(* CODESYS project Example10_PLC.project

Project tree, tasks and I/O mapping:
  Device : CODESYS Control Win V3, 3S - Smart Software Solutions GmbH, order no. 305021, version 3.5.7.0
    application Application
      libraries: Standard, * (System)
      task MainTask (cyclic, interval t#20ms, priority 1) calls PLC_PRG
      program PLC_PRG [ST]
      global variables GVL
      function block FB_G4LTL [ST]
    Ethernet : Ethernet, 3S - Smart Software Solutions GmbH, version 3.5.7.0
      Modbus_TCP_Master : Modbus TCP Master, 3S - Smart Software Solutions GmbH, version 3.5.6.0
          settings: AutoReconnect = TRUE
        Modbus_TCP_Slave : Modbus TCP Slave, 3S - Smart Software Solutions GmbH, version 3.5.7.0
            settings: Unit-ID = 1; IPAddress = [127, 0, 0, 1]; Channel 0.Function Code = 4; Channel 0.Read Offset = 16#0000; Channel 0.Read Length = 1; Channel 0.Write Offset = 0; Channel 0.Write Length = 0; Channel 0.Cycle Time = 100; Channel 1.Function Code = 4; Channel 1.Read Offset = 16#0001; Channel 1.Read Length = 1; Channel 1.Write Offset = 0; Channel 1.Write Length = 0; Channel 1.Cycle Time = 100; Channel 2.Function Code = 4; Channel 2.Read Offset = 16#0002; Channel 2.Read Length = 1; Channel 2.Write Offset = 0; Channel 2.Write Length = 0; Channel 2.Cycle Time = 100; Channel 3.Function Code = 4; Channel 3.Read Offset = 16#0003; Channel 3.Read Length = 1; Channel 3.Write Offset = 0; Channel 3.Write Length = 0; Channel 3.Cycle Time = 100; Channel 4.Function Code = 4; Channel 4.Read Offset = 16#0004; Channel 4.Read Length = 1; Channel 4.Write Offset = 0; Channel 4.Write Length = 0; Channel 4.Cycle Time = 100; Channel 5.Function Code = 6; Channel 5.Read Offset = 0; Channel 5.Read Length = 0; Channel 5.Write Offset = 16#0000; Channel 5.Write Length = 1; Channel 5.Cycle Time = 100; Channel 6.Function Code = 6; Channel 6.Read Offset = 0;
              Channel 6.Read Length = 0; Channel 6.Write Offset = 16#0002; Channel 6.Write Length = 1; Channel 6.Cycle Time = 100; Channel 7.Function Code = 6; Channel 7.Read Offset = 0; Channel 7.Read Length = 0; Channel 7.Write Offset = 16#0003; Channel 7.Write Length = 1; Channel 7.Cycle Time = 100; Channel 8.Function Code = 6; Channel 8.Read Offset = 0; Channel 8.Read Length = 0; Channel 8.Write Offset = 16#0004; Channel 8.Write Length = 1; Channel 8.Cycle Time = 100; Channel 9.Function Code = 6; Channel 9.Read Offset = 0; Channel 9.Read Length = 0; Channel 9.Write Offset = 16#0001; Channel 9.Write Length = 1; Channel 9.Cycle Time = 100
            input  Application.dIn0 : BOOL  // Channel 0.Channel 0.Bit0
            input  Application.dIn1 : BOOL  // Channel 1.Channel 1.Bit0
            input  Application.dIn2 : BOOL  // Channel 2.Channel 2.Bit0
            input  Application.dIn3 : BOOL  // Channel 3.Channel 3.Bit0
            input  Application.dIn4 : BOOL  // Channel 4.Channel 4.Bit0
            output Application.dOut0 : BOOL  // Channel 5.Channel 5.Bit0
            output Application.dOut2 : BOOL  // Channel 6.Channel 6.Bit0
            output Application.dOut3 : BOOL  // Channel 7.Channel 7.Bit0
            output Application.dOut4 : BOOL  // Channel 8.Channel 8.Bit0
            output Application.dOut1 : BOOL  // Channel 9.Channel 9.Bit0
            unmapped channels: Channel 0, Channel 1, Channel 2, Channel 3, Channel 4, Channel 5, Channel 6, Channel 7, Channel 8, Channel 9
*)

// Device/Application/GVL
VAR_GLOBAL
	
dIn0 : BOOL;
dIn1 : BOOL;
dIn2 : BOOL;
dIn3 : BOOL;
dIn4 : BOOL;

dOut0 : BOOL;
dOut1 : BOOL; 
dOut2 : BOOL; 
dOut3 : BOOL; 
dOut4 : BOOL; 
END_VAR

// Device/Application/PLC_PRG
PROGRAM PLC_PRG


VAR 
	fb: FB_G4LTL;

END_VAR

// Direct looping
// Assign pins (from global variable to function block) 
fb.x0 := dIn0;
fb.x1 := dIn1;
fb.x2 := dIn2;
fb.x3 := dIn3;
fb.x10 := dIn4;

// Assign pins (from function block to global variable)
dOut0 := fb.y0;
dOut1 := fb.y1;
dOut2 := fb.y2;
dOut3 := fb.y3;

// Run the function block
fb();

END_PROGRAM

// Device/Application/FB_G4LTL
FUNCTION_BLOCK FB_G4LTL

   (* Variable definition *)
   VAR_INPUT
      x0	: BOOL;
      x1	: BOOL;
      x2	: BOOL;
      x3	: BOOL;
      x10	: BOOL;
   END_VAR
   VAR_OUTPUT
      y0	: BOOL;
      y1	: BOOL;
      y2	: BOOL;
      y3	: BOOL;
   END_VAR
   VAR
   (* Control logic for y0, y1; the total number of states equals to 13 *)
      cstate23	: LINT := 0;
   (* Control logic for y2, y3; the total number of states equals to 37 *)
      cstate64	: LINT := 0;  
	  
      t0	: TON;
      t0_reset	: BOOL := FALSE;
      t0_up	: BOOL := FALSE;
      t0_start	: BOOL := FALSE;
      t1	: TON;
      t1_reset	: BOOL := FALSE;
      t1_up	: BOOL := FALSE;
      t1_start	: BOOL := FALSE;
	  
      T0_VALUE	: TIME := TIME#3S;
      T1_VALUE	: TIME := TIME#6S;	  
   END_VAR

   (* Constant definition  *)

    (* Control logic for y0, y1*)
CASE cstate23 OF
262:
    IF ((x0 = TRUE) AND  (x1 = FALSE) AND  ( TRUE ) AND  (x10 = TRUE)) OR ((x0 = TRUE) AND  (x1 = TRUE) AND  (x2 = FALSE) AND  (x10 = TRUE)) OR ((x0 = TRUE) AND  (x1 = TRUE) AND  (x2 = TRUE) AND  ( TRUE )) THEN 
        cstate23 := 27; y0 := FALSE; y1 := FALSE;  
    ELSIF ((x0 = FALSE) AND  (x1 = FALSE) AND  ( TRUE ) AND  (x10 = TRUE)) OR ((x0 = FALSE) AND  (x1 = TRUE) AND  (x2 = FALSE) AND  (x10 = TRUE)) OR ((x0 = FALSE) AND  (x1 = TRUE) AND  (x2 = TRUE) AND  ( TRUE )) THEN 
        cstate23 := 20; y0 := FALSE; y1 := FALSE;  
    ELSIF ((x0 = FALSE) AND  (x1 = FALSE) AND  ( TRUE ) AND  (x10 = FALSE)) THEN 
        cstate23 := 20; y0 := TRUE; y1 := FALSE;  
    ELSIF ((x0 = TRUE) AND  (x1 = TRUE) AND  (x2 = FALSE) AND  (x10 = FALSE)) THEN 
        cstate23 := 265; y0 := FALSE; y1 := TRUE;  
    ELSIF ((x0 = TRUE) AND  (x1 = FALSE) AND  ( TRUE ) AND  (x10 = FALSE)) THEN 
        cstate23 := 262; y0 := TRUE; y1 := FALSE;  
    ELSIF ((x0 = FALSE) AND  (x1 = TRUE) AND  (x2 = FALSE) AND  (x10 = FALSE)) THEN 
        cstate23 := 260; y0 := FALSE; y1 := TRUE;  
    END_IF;
669:
    IF ((x0 = TRUE) AND  (x1 = FALSE) AND  ( TRUE ) AND  (x10 = TRUE)) OR ((x0 = TRUE) AND  (x1 = TRUE) AND  (x2 = FALSE) AND  (x10 = TRUE)) OR ((x0 = TRUE) AND  (x1 = TRUE) AND  (x2 = TRUE) AND  ( TRUE )) THEN 
        cstate23 := 27; y0 := FALSE; y1 := FALSE;  
    ELSIF ((x0 = FALSE) AND  (x1 = FALSE) AND  ( TRUE ) AND  (x10 = TRUE)) OR ((x0 = FALSE) AND  (x1 = TRUE) AND  (x2 = FALSE) AND  (x10 = TRUE)) OR ((x0 = FALSE) AND  (x1 = TRUE) AND  (x2 = TRUE) AND  ( TRUE )) THEN 
        cstate23 := 20; y0 := FALSE; y1 := FALSE;  
    ELSIF ((x0 = FALSE) AND  ( TRUE ) AND  (x2 = FALSE) AND  (x10 = FALSE)) THEN 
        cstate23 := 260; y0 := FALSE; y1 := TRUE;  
    ELSIF ((x0 = TRUE) AND  (x1 = TRUE) AND  (x2 = FALSE) AND  (x10 = FALSE)) THEN 
        cstate23 := 265; y0 := FALSE; y1 := TRUE;  
    ELSIF ((x0 = FALSE) AND  (x1 = FALSE) AND  (x2 = TRUE) AND  (x10 = FALSE)) THEN 
        cstate23 := 20; y0 := TRUE; y1 := FALSE;  
    ELSIF ((x0 = TRUE) AND  (x1 = FALSE) AND  (x2 = TRUE) AND  (x10 = FALSE)) THEN 
        cstate23 := 262; y0 := TRUE; y1 := FALSE;  
    ELSIF ((x0 = TRUE) AND  (x1 = FALSE) AND  (x2 = FALSE) AND  (x10 = FALSE)) THEN 
        cstate23 := 669; y0 := TRUE; y1 := TRUE;  
    END_IF;
260:
    IF ((x0 = TRUE) AND  (x1 = FALSE) AND  ( TRUE ) AND  (x10 = TRUE)) OR ((x0 = TRUE) AND  (x1 = TRUE) AND  (x2 = FALSE) AND  (x10 = TRUE)) OR ((x0 = TRUE) AND  (x1 = TRUE) AND  (x2 = TRUE) AND  ( TRUE )) THEN 
        cstate23 := 27; y0 := FALSE; y1 := FALSE;  
    ELSIF ((x0 = FALSE) AND  ( TRUE ) AND  (x2 = FALSE) AND  (x10 = TRUE)) OR ((x0 = FALSE) AND  ( TRUE ) AND  (x2 = TRUE) AND  ( TRUE )) THEN 
        cstate23 := 20; y0 := FALSE; y1 := FALSE;  
    ELSIF ((x0 = FALSE) AND  ( TRUE ) AND  (x2 = FALSE) AND  (x10 = FALSE)) THEN 
        cstate23 := 260; y0 := FALSE; y1 := TRUE;  
    ELSIF ((x0 = TRUE) AND  (x1 = TRUE) AND  (x2 = FALSE) AND  (x10 = FALSE)) THEN 
        cstate23 := 265; y0 := FALSE; y1 := TRUE;  
    ELSIF ((x0 = TRUE) AND  (x1 = FALSE) AND  (x2 = TRUE) AND  (x10 = FALSE)) THEN 
        cstate23 := 262; y0 := TRUE; y1 := FALSE;  
    ELSIF ((x0 = TRUE) AND  (x1 = FALSE) AND  (x2 = FALSE) AND  (x10 = FALSE)) THEN 
        cstate23 := 669; y0 := TRUE; y1 := TRUE;  
    END_IF;
18:
    IF ((x0 = TRUE) AND  ( TRUE ) AND  ( TRUE ) AND  (x10 = TRUE)) THEN 
        cstate23 := 27; y0 := FALSE; y1 := FALSE;  
    ELSIF ((x0 = FALSE) AND  ( TRUE ) AND  ( TRUE ) AND  (x10 = TRUE)) THEN 
        cstate23 := 20; y0 := FALSE; y1 := FALSE;  
    ELSIF ((x0 = FALSE) AND  (x1 = FALSE) AND  ( TRUE ) AND  (x10 = FALSE)) OR ((x0 = FALSE) AND  (x1 = TRUE) AND  (x2 = TRUE) AND  (x10 = FALSE)) THEN 
        cstate23 := 18; y0 := FALSE; y1 := FALSE;  
    ELSIF ((x0 = TRUE) AND  (x1 = TRUE) AND  (x2 = FALSE) AND  (x10 = FALSE)) THEN 
        cstate23 := 31; y0 := FALSE; y1 := TRUE;  
    ELSIF ((x0 = TRUE) AND  (x1 = TRUE) AND  (x2 = TRUE) AND  (x10 = FALSE)) THEN 
        cstate23 := 25; y0 := FALSE; y1 := FALSE;  
    ELSIF ((x0 = TRUE) AND  (x1 = FALSE) AND  ( TRUE ) AND  (x10 = FALSE)) THEN 
        cstate23 := 257; y0 := TRUE; y1 := FALSE;  
    ELSIF ((x0 = FALSE) AND  (x1 = TRUE) AND  (x2 = FALSE) AND  (x10 = FALSE)) THEN 
        cstate23 := 24; y0 := FALSE; y1 := TRUE;  
    END_IF;
24:
    IF ((x0 = TRUE) AND  ( TRUE ) AND  ( TRUE ) AND  (x10 = TRUE)) THEN 
        cstate23 := 27; y0 := FALSE; y1 := FALSE;  
    ELSIF ((x0 = FALSE) AND  ( TRUE ) AND  ( TRUE ) AND  (x10 = TRUE)) THEN 
        cstate23 := 20; y0 := FALSE; y1 := FALSE;  
    ELSIF ((x0 = FALSE) AND  ( TRUE ) AND  (x2 = FALSE) AND  (x10 = FALSE)) THEN 
        cstate23 := 24; y0 := FALSE; y1 := TRUE;  
    ELSIF ((x0 = TRUE) AND  (x1 = TRUE) AND  (x2 = FALSE) AND  (x10 = FALSE)) THEN 
        cstate23 := 31; y0 := FALSE; y1 := TRUE;  
    ELSIF ((x0 = TRUE) AND  (x1 = TRUE) AND  (x2 = TRUE) AND  (x10 = FALSE)) THEN 
        cstate23 := 25; y0 := FALSE; y1 := FALSE;  
    ELSIF ((x0 = FALSE) AND  ( TRUE ) AND  (x2 = TRUE) AND  (x10 = FALSE)) THEN 
        cstate23 := 18; y0 := FALSE; y1 := FALSE;  
    ELSIF ((x0 = TRUE) AND  (x1 = FALSE) AND  (x2 = TRUE) AND  (x10 = FALSE)) THEN 
        cstate23 := 257; y0 := TRUE; y1 := FALSE;  
    ELSIF ((x0 = TRUE) AND  (x1 = FALSE) AND  (x2 = FALSE) AND  (x10 = FALSE)) THEN 
        cstate23 := 279; y0 := TRUE; y1 := TRUE;  
    END_IF;
25:
    IF ((x0 = TRUE) AND  ( TRUE ) AND  ( TRUE ) AND  (x10 = TRUE)) THEN 
        cstate23 := 27; y0 := FALSE; y1 := FALSE;  
    ELSIF ((x0 = FALSE) AND  ( TRUE ) AND  ( TRUE ) AND  (x10 = TRUE)) THEN 
        cstate23 := 20; y0 := FALSE; y1 := FALSE;  
    ELSIF ((x0 = FALSE) AND  (x1 = FALSE) AND  ( TRUE ) AND  (x10 = FALSE)) THEN 
        cstate23 := 18; y0 := TRUE; y1 := FALSE;  
    ELSIF ((x0 = TRUE) AND  (x1 = TRUE) AND  (x2 = FALSE) AND  (x10 = FALSE)) THEN 
        cstate23 := 31; y0 := FALSE; y1 := TRUE;  
    ELSIF ((x0 = TRUE) AND  (x1 = TRUE) AND  (x2 = TRUE) AND  (x10 = FALSE)) THEN 
        cstate23 := 25; y0 := FALSE; y1 := FALSE;  
    ELSIF ((x0 = FALSE) AND  (x1 = TRUE) AND  (x2 = TRUE) AND  (x10 = FALSE)) THEN 
        cstate23 := 18; y0 := FALSE; y1 := FALSE;  
    ELSIF ((x0 = TRUE) AND  (x1 = FALSE) AND  ( TRUE ) AND  (x10 = FALSE)) THEN 
        cstate23 := 25; y0 := TRUE; y1 := FALSE;  
    ELSIF ((x0 = FALSE) AND  (x1 = TRUE) AND  (x2 = FALSE) AND  (x10 = FALSE)) THEN 
        cstate23 := 24; y0 := FALSE; y1 := TRUE;  
    END_IF;
27:
    IF ((x0 = TRUE) AND  (x1 = FALSE) AND  ( TRUE ) AND  (x10 = TRUE)) OR ((x0 = TRUE) AND  (x1 = TRUE) AND  (x2 = FALSE) AND  (x10 = TRUE)) OR ((x0 = TRUE) AND  (x1 = TRUE) AND  (x2 = TRUE) AND  ( TRUE )) THEN 
        cstate23 := 27; y0 := FALSE; y1 := FALSE;  
    ELSIF ((x0 = FALSE) AND  (x1 = FALSE) AND  ( TRUE ) AND  (x10 = TRUE)) OR ((x0 = FALSE) AND  (x1 = TRUE) AND  (x2 = FALSE) AND  (x10 = TRUE)) OR ((x0 = FALSE) AND  (x1 = TRUE) AND  (x2 = TRUE) AND  ( TRUE )) THEN 
        cstate23 := 20; y0 := FALSE; y1 := FALSE;  
    ELSIF ((x0 = FALSE) AND  (x1 = FALSE) AND  ( TRUE ) AND  (x10 = FALSE)) THEN 
        cstate23 := 20; y0 := TRUE; y1 := FALSE;  
    ELSIF ((x0 = TRUE) AND  (x1 = TRUE) AND  (x2 = FALSE) AND  (x10 = FALSE)) THEN 
        cstate23 := 265; y0 := FALSE; y1 := TRUE;  
    ELSIF ((x0 = TRUE) AND  (x1 = FALSE) AND  ( TRUE ) AND  (x10 = FALSE)) THEN 
        cstate23 := 27; y0 := TRUE; y1 := FALSE;  
    ELSIF ((x0 = FALSE) AND  (x1 = TRUE) AND  (x2 = FALSE) AND  (x10 = FALSE)) THEN 
        cstate23 := 260; y0 := FALSE; y1 := TRUE;  
    END_IF;
20:
    IF ((x0 = TRUE) AND  (x1 = FALSE) AND  ( TRUE ) AND  (x10 = TRUE)) OR ((x0 = TRUE) AND  (x1 = TRUE) AND  (x2 = FALSE) AND  (x10 = TRUE)) OR ((x0 = TRUE) AND  (x1 = TRUE) AND  (x2 = TRUE) AND  ( TRUE )) THEN 
        cstate23 := 27; y0 := FALSE; y1 := FALSE;  
    ELSIF ((x0 = FALSE) AND  (x1 = FALSE) AND  ( TRUE ) AND  ( TRUE )) OR ((x0 = FALSE) AND  (x1 = TRUE) AND  (x2 = FALSE) AND  (x10 = TRUE)) OR ((x0 = FALSE) AND  (x1 = TRUE) AND  (x2 = TRUE) AND  ( TRUE )) THEN 
        cstate23 := 20; y0 := FALSE; y1 := FALSE;  
    ELSIF ((x0 = TRUE) AND  (x1 = TRUE) AND  (x2 = FALSE) AND  (x10 = FALSE)) THEN 
        cstate23 := 265; y0 := FALSE; y1 := TRUE;  
    ELSIF ((x0 = TRUE) AND  (x1 = FALSE) AND  ( TRUE ) AND  (x10 = FALSE)) THEN 
        cstate23 := 262; y0 := TRUE; y1 := FALSE;  
    ELSIF ((x0 = FALSE) AND  (x1 = TRUE) AND  (x2 = FALSE) AND  (x10 = FALSE)) THEN 
        cstate23 := 260; y0 := FALSE; y1 := TRUE;  
    END_IF;
0:
    IF ((x0 = TRUE) AND  ( TRUE ) AND  ( TRUE ) AND  (x10 = TRUE)) THEN 
        cstate23 := 27; y0 := FALSE; y1 := FALSE;  
    ELSIF ((x0 = FALSE) AND  ( TRUE ) AND  ( TRUE ) AND  (x10 = TRUE)) THEN 
        cstate23 := 20; y0 := FALSE; y1 := FALSE;  
    ELSIF ((x0 = FALSE) AND  (x1 = FALSE) AND  ( TRUE ) AND  (x10 = FALSE)) OR ((x0 = FALSE) AND  (x1 = TRUE) AND  (x2 = TRUE) AND  (x10 = FALSE)) THEN 
        cstate23 := 18; y0 := FALSE; y1 := FALSE;  
    ELSIF ((x0 = TRUE) AND  (x1 = TRUE) AND  (x2 = FALSE) AND  (x10 = FALSE)) THEN 
        cstate23 := 31; y0 := FALSE; y1 := TRUE;  
    ELSIF ((x0 = TRUE) AND  (x1 = FALSE) AND  ( TRUE ) AND  (x10 = FALSE)) OR ((x0 = TRUE) AND  (x1 = TRUE) AND  (x2 = TRUE) AND  (x10 = FALSE)) THEN 
        cstate23 := 25; y0 := FALSE; y1 := FALSE;  
    ELSIF ((x0 = FALSE) AND  (x1 = TRUE) AND  (x2 = FALSE) AND  (x10 = FALSE)) THEN 
        cstate23 := 24; y0 := FALSE; y1 := TRUE;  
    END_IF;
279:
    IF ((x0 = TRUE) AND  ( TRUE ) AND  ( TRUE ) AND  (x10 = TRUE)) THEN 
        cstate23 := 27; y0 := FALSE; y1 := FALSE;  
    ELSIF ((x0 = FALSE) AND  ( TRUE ) AND  ( TRUE ) AND  (x10 = TRUE)) THEN 
        cstate23 := 20; y0 := FALSE; y1 := FALSE;  
    ELSIF ((x0 = FALSE) AND  ( TRUE ) AND  (x2 = FALSE) AND  (x10 = FALSE)) THEN 
        cstate23 := 24; y0 := FALSE; y1 := TRUE;  
    ELSIF ((x0 = TRUE) AND  (x1 = TRUE) AND  (x2 = FALSE) AND  (x10 = FALSE)) THEN 
        cstate23 := 31; y0 := FALSE; y1 := TRUE;  
    ELSIF ((x0 = TRUE) AND  (x1 = TRUE) AND  (x2 = TRUE) AND  (x10 = FALSE)) THEN 
        cstate23 := 25; y0 := FALSE; y1 := FALSE;  
    ELSIF ((x0 = FALSE) AND  (x1 = FALSE) AND  (x2 = TRUE) AND  (x10 = FALSE)) THEN 
        cstate23 := 18; y0 := TRUE; y1 := FALSE;  
    ELSIF ((x0 = FALSE) AND  (x1 = TRUE) AND  (x2 = TRUE) AND  (x10 = FALSE)) THEN 
        cstate23 := 18; y0 := FALSE; y1 := FALSE;  
    ELSIF ((x0 = TRUE) AND  (x1 = FALSE) AND  (x2 = TRUE) AND  (x10 = FALSE)) THEN 
        cstate23 := 257; y0 := TRUE; y1 := FALSE;  
    ELSIF ((x0 = TRUE) AND  (x1 = FALSE) AND  (x2 = FALSE) AND  (x10 = FALSE)) THEN 
        cstate23 := 279; y0 := TRUE; y1 := TRUE;  
    END_IF;
31:
    IF ((x0 = TRUE) AND  ( TRUE ) AND  ( TRUE ) AND  (x10 = TRUE)) THEN 
        cstate23 := 27; y0 := FALSE; y1 := FALSE;  
    ELSIF ((x0 = FALSE) AND  ( TRUE ) AND  ( TRUE ) AND  (x10 = TRUE)) THEN 
        cstate23 := 20; y0 := FALSE; y1 := FALSE;  
    ELSIF ((x0 = FALSE) AND  ( TRUE ) AND  (x2 = FALSE) AND  (x10 = FALSE)) THEN 
        cstate23 := 24; y0 := FALSE; y1 := TRUE;  
    ELSIF ((x0 = TRUE) AND  ( TRUE ) AND  (x2 = FALSE) AND  (x10 = FALSE)) THEN 
        cstate23 := 31; y0 := FALSE; y1 := TRUE;  
    ELSIF ((x0 = TRUE) AND  (x1 = TRUE) AND  (x2 = TRUE) AND  (x10 = FALSE)) THEN 
        cstate23 := 25; y0 := FALSE; y1 := FALSE;  
    ELSIF ((x0 = FALSE) AND  (x1 = FALSE) AND  (x2 = TRUE) AND  (x10 = FALSE)) THEN 
        cstate23 := 18; y0 := TRUE; y1 := FALSE;  
    ELSIF ((x0 = FALSE) AND  (x1 = TRUE) AND  (x2 = TRUE) AND  (x10 = FALSE)) THEN 
        cstate23 := 18; y0 := FALSE; y1 := FALSE;  
    ELSIF ((x0 = TRUE) AND  (x1 = FALSE) AND  (x2 = TRUE) AND  (x10 = FALSE)) THEN 
        cstate23 := 25; y0 := TRUE; y1 := FALSE;  
    END_IF;
257:
    IF ((x0 = TRUE) AND  ( TRUE ) AND  ( TRUE ) AND  (x10 = TRUE)) THEN 
        cstate23 := 27; y0 := FALSE; y1 := FALSE;  
    ELSIF ((x0 = FALSE) AND  ( TRUE ) AND  ( TRUE ) AND  (x10 = TRUE)) THEN 
        cstate23 := 20; y0 := FALSE; y1 := FALSE;  
    ELSIF ((x0 = FALSE) AND  (x1 = FALSE) AND  ( TRUE ) AND  (x10 = FALSE)) THEN 
        cstate23 := 18; y0 := TRUE; y1 := FALSE;  
    ELSIF ((x0 = TRUE) AND  (x1 = TRUE) AND  (x2 = FALSE) AND  (x10 = FALSE)) THEN 
        cstate23 := 31; y0 := FALSE; y1 := TRUE;  
    ELSIF ((x0 = TRUE) AND  (x1 = TRUE) AND  (x2 = TRUE) AND  (x10 = FALSE)) THEN 
        cstate23 := 25; y0 := FALSE; y1 := FALSE;  
    ELSIF ((x0 = FALSE) AND  (x1 = TRUE) AND  (x2 = TRUE) AND  (x10 = FALSE)) THEN 
        cstate23 := 18; y0 := FALSE; y1 := FALSE;  
    ELSIF ((x0 = TRUE) AND  (x1 = FALSE) AND  ( TRUE ) AND  (x10 = FALSE)) THEN 
        cstate23 := 257; y0 := TRUE; y1 := FALSE;  
    ELSIF ((x0 = FALSE) AND  (x1 = TRUE) AND  (x2 = FALSE) AND  (x10 = FALSE)) THEN 
        cstate23 := 24; y0 := FALSE; y1 := TRUE;  
    END_IF;
265:
    IF ((x0 = TRUE) AND  (x1 = FALSE) AND  ( TRUE ) AND  (x10 = TRUE)) OR ((x0 = TRUE) AND  (x1 = TRUE) AND  (x2 = FALSE) AND  (x10 = TRUE)) OR ((x0 = TRUE) AND  (x1 = TRUE) AND  (x2 = TRUE) AND  ( TRUE )) THEN 
        cstate23 := 27; y0 := FALSE; y1 := FALSE;  
    ELSIF ((x0 = FALSE) AND  (x1 = FALSE) AND  ( TRUE ) AND  (x10 = TRUE)) OR ((x0 = FALSE) AND  (x1 = TRUE) AND  (x2 = FALSE) AND  (x10 = TRUE)) OR ((x0 = FALSE) AND  (x1 = TRUE) AND  (x2 = TRUE) AND  ( TRUE )) THEN 
        cstate23 := 20; y0 := FALSE; y1 := FALSE;  
    ELSIF ((x0 = FALSE) AND  ( TRUE ) AND  (x2 = FALSE) AND  (x10 = FALSE)) THEN 
        cstate23 := 260; y0 := FALSE; y1 := TRUE;  
    ELSIF ((x0 = TRUE) AND  ( TRUE ) AND  (x2 = FALSE) AND  (x10 = FALSE)) THEN 
        cstate23 := 265; y0 := FALSE; y1 := TRUE;  
    ELSIF ((x0 = FALSE) AND  (x1 = FALSE) AND  (x2 = TRUE) AND  (x10 = FALSE)) THEN 
        cstate23 := 20; y0 := TRUE; y1 := FALSE;  
    ELSIF ((x0 = TRUE) AND  (x1 = FALSE) AND  (x2 = TRUE) AND  (x10 = FALSE)) THEN 
        cstate23 := 27; y0 := TRUE; y1 := FALSE;  
    END_IF;
END_CASE;


 (* Control logic *)
CASE cstate64 OF
19:
    IF ((x2 = FALSE) AND  ( TRUE ) AND  ( TRUE ) AND  (t0.Q = FALSE) AND  (t1.Q = FALSE)) THEN 
        cstate64 := 19; y2 := FALSE; y3 := FALSE; t0_start := FALSE;t1_start := FALSE; 
    ELSIF ((x2 = FALSE) AND  ( TRUE ) AND  (x10 = FALSE) AND  (t0.Q = FALSE) AND  (t1.Q = TRUE)) THEN 
        cstate64 := 20; y2 := FALSE; y3 := FALSE; t0_start := FALSE;t1_start := FALSE; 
    ELSIF ((x2 = FALSE) AND  ( TRUE ) AND  (x10 = FALSE) AND  (t0.Q = TRUE) AND  ( TRUE )) THEN 
        cstate64 := 37; y2 := FALSE; y3 := TRUE; t0_start := FALSE;t1_start := TRUE; t1_up := FALSE; 
    ELSIF ((x2 = FALSE) AND  ( TRUE ) AND  (x10 = TRUE) AND  (t0.Q = FALSE) AND  (t1.Q = TRUE)) THEN 
        cstate64 := 20; y2 := FALSE; y3 := FALSE; t0_start := FALSE;t1_start := FALSE; 
    ELSIF ((x2 = FALSE) AND  ( TRUE ) AND  (x10 = TRUE) AND  (t0.Q = TRUE) AND  (t1.Q = FALSE)) THEN 
        cstate64 := 34; y2 := FALSE; y3 := FALSE; t0_start := FALSE;t1_start := FALSE; 
    ELSIF ((x2 = FALSE) AND  ( TRUE ) AND  (x10 = TRUE) AND  (t0.Q = TRUE) AND  (t1.Q = TRUE)) THEN 
        cstate64 := 33; y2 := FALSE; y3 := FALSE; t0_start := FALSE;t1_start := FALSE; 
    ELSIF ((x2 = TRUE) AND  ( TRUE ) AND  (x10 = FALSE) AND  (t0.Q = FALSE) AND  (t1.Q = FALSE)) THEN 
        cstate64 := 83; y2 := TRUE; y3 := FALSE; t0_start := TRUE; t0_up := FALSE;t1_start := FALSE; 
    ELSIF ((x2 = TRUE) AND  ( TRUE ) AND  (x10 = FALSE) AND  (t0.Q = FALSE) AND  (t1.Q = TRUE)) THEN 
        cstate64 := 84; y2 := TRUE; y3 := FALSE; t0_start := TRUE; t0_up := FALSE;t1_start := FALSE; 
    ELSIF ((x2 = TRUE) AND  ( TRUE ) AND  (x10 = FALSE) AND  (t0.Q = TRUE) AND  ( TRUE )) THEN 
        cstate64 := 86; y2 := TRUE; y3 := TRUE; t0_start := TRUE; t0_up := FALSE;t1_start := TRUE; t1_up := FALSE; 
    ELSIF ((x2 = TRUE) AND  ( TRUE ) AND  (x10 = TRUE) AND  (t0.Q = FALSE) AND  (t1.Q = FALSE)) THEN 
        cstate64 := 51; y2 := FALSE; y3 := FALSE; t0_start := FALSE;t1_start := FALSE; 
    ELSIF ((x2 = TRUE) AND  ( TRUE ) AND  (x10 = TRUE) AND  (t0.Q = FALSE) AND  (t1.Q = TRUE)) THEN 
        cstate64 := 52; y2 := FALSE; y3 := FALSE; t0_start := FALSE;t1_start := FALSE; 
    ELSIF ((x2 = TRUE) AND  ( TRUE ) AND  (x10 = TRUE) AND  (t0.Q = TRUE) AND  (t1.Q = FALSE)) THEN 
        cstate64 := 66; y2 := FALSE; y3 := FALSE; t0_start := FALSE;t1_start := FALSE; 
    ELSIF ((x2 = TRUE) AND  ( TRUE ) AND  (x10 = TRUE) AND  (t0.Q = TRUE) AND  (t1.Q = TRUE)) THEN 
        cstate64 := 65; y2 := FALSE; y3 := FALSE; t0_start := FALSE;t1_start := FALSE; 
    END_IF;
35:
    IF ((x2 = FALSE) AND  ( TRUE ) AND  ( TRUE ) AND  (t0.Q = FALSE) AND  (t1.Q = FALSE)) THEN 
        cstate64 := 35; y2 := FALSE; y3 := FALSE; t0_start := FALSE;t1_start := FALSE; 
    ELSIF ((x2 = FALSE) AND  ( TRUE ) AND  (x10 = FALSE) AND  (t0.Q = FALSE) AND  (t1.Q = TRUE)) THEN 
        cstate64 := 36; y2 := FALSE; y3 := FALSE; t0_start := FALSE;t1_start := FALSE; 
    ELSIF ((x2 = FALSE) AND  ( TRUE ) AND  (x10 = FALSE) AND  (t0.Q = TRUE) AND  ( TRUE )) THEN 
        cstate64 := 37; y2 := FALSE; y3 := TRUE; t0_start := FALSE;t1_start := TRUE; t1_up := FALSE; 
    ELSIF ((x2 = FALSE) AND  ( TRUE ) AND  (x10 = TRUE) AND  (t0.Q = FALSE) AND  (t1.Q = TRUE)) THEN 
        cstate64 := 36; y2 := FALSE; y3 := FALSE; t0_start := FALSE;t1_start := FALSE; 
    ELSIF ((x2 = FALSE) AND  ( TRUE ) AND  (x10 = TRUE) AND  (t0.Q = TRUE) AND  (t1.Q = FALSE)) THEN 
        cstate64 := 34; y2 := FALSE; y3 := FALSE; t0_start := FALSE;t1_start := FALSE; 
    ELSIF ((x2 = FALSE) AND  ( TRUE ) AND  (x10 = TRUE) AND  (t0.Q = TRUE) AND  (t1.Q = TRUE)) THEN 
        cstate64 := 33; y2 := FALSE; y3 := FALSE; t0_start := FALSE;t1_start := FALSE; 
    ELSIF ((x2 = TRUE) AND  ( TRUE ) AND  (x10 = FALSE) AND  (t0.Q = FALSE) AND  (t1.Q = FALSE)) THEN 
        cstate64 := 83; y2 := TRUE; y3 := FALSE; t0_start := TRUE; t0_up := FALSE;t1_start := FALSE; 
    ELSIF ((x2 = TRUE) AND  ( TRUE ) AND  (x10 = FALSE) AND  (t0.Q = FALSE) AND  (t1.Q = TRUE)) THEN 
        cstate64 := 84; y2 := TRUE; y3 := FALSE; t0_start := TRUE; t0_up := FALSE;t1_start := FALSE; 
    ELSIF ((x2 = TRUE) AND  ( TRUE ) AND  (x10 = FALSE) AND  (t0.Q = TRUE) AND  ( TRUE )) THEN 
        cstate64 := 86; y2 := TRUE; y3 := TRUE; t0_start := TRUE; t0_up := FALSE;t1_start := TRUE; t1_up := FALSE; 
    ELSIF ((x2 = TRUE) AND  ( TRUE ) AND  (x10 = TRUE) AND  (t0.Q = FALSE) AND  (t1.Q = FALSE)) THEN 
        cstate64 := 67; y2 := FALSE; y3 := FALSE; t0_start := FALSE;t1_start := FALSE; 
    ELSIF ((x2 = TRUE) AND  ( TRUE ) AND  (x10 = TRUE) AND  (t0.Q = FALSE) AND  (t1.Q = TRUE)) THEN 
        cstate64 := 68; y2 := FALSE; y3 := FALSE; t0_start := FALSE;t1_start := FALSE; 
    ELSIF ((x2 = TRUE) AND  ( TRUE ) AND  (x10 = TRUE) AND  (t0.Q = TRUE) AND  (t1.Q = FALSE)) THEN 
        cstate64 := 66; y2 := FALSE; y3 := FALSE; t0_start := FALSE;t1_start := FALSE; 
    ELSIF ((x2 = TRUE) AND  ( TRUE ) AND  (x10 = TRUE) AND  (t0.Q = TRUE) AND  (t1.Q = TRUE)) THEN 
        cstate64 := 65; y2 := FALSE; y3 := FALSE; t0_start := FALSE;t1_start := FALSE; 
    END_IF;
36:
    IF ((x2 = FALSE) AND  ( TRUE ) AND  (x10 = FALSE) AND  (t0.Q = FALSE) AND  (t1.Q = FALSE)) OR ((x2 = FALSE) AND  ( TRUE ) AND  (x10 = TRUE) AND  (t0.Q = FALSE) AND  ( TRUE )) THEN 
        cstate64 := 36; y2 := FALSE; y3 := FALSE; t0_start := FALSE;t1_start := FALSE; 
    ELSIF ((x2 = FALSE) AND  ( TRUE ) AND  (x10 = FALSE) AND  (t0.Q = FALSE) AND  (t1.Q = TRUE)) THEN 
        cstate64 := 36; y2 := FALSE; y3 := FALSE; t0_start := FALSE;t1_start := FALSE; 
    ELSIF ((x2 = FALSE) AND  ( TRUE ) AND  (x10 = FALSE) AND  (t0.Q = TRUE) AND  ( TRUE )) THEN 
        cstate64 := 40; y2 := FALSE; y3 := TRUE; t0_start := FALSE;t1_start := TRUE; t1_up := FALSE; 
    ELSIF ((x2 = FALSE) AND  ( TRUE ) AND  (x10 = TRUE) AND  (t0.Q = TRUE) AND  ( TRUE )) THEN 
        cstate64 := 33; y2 := FALSE; y3 := FALSE; t0_start := FALSE;t1_start := FALSE; 
    ELSIF ((x2 = TRUE) AND  ( TRUE ) AND  (x10 = FALSE) AND  (t0.Q = FALSE) AND  (t1.Q = FALSE)) THEN 
        cstate64 := 84; y2 := TRUE; y3 := FALSE; t0_start := TRUE; t0_up := FALSE;t1_start := FALSE; 
    ELSIF ((x2 = TRUE) AND  ( TRUE ) AND  (x10 = FALSE) AND  (t0.Q = FALSE) AND  (t1.Q = TRUE)) THEN 
        cstate64 := 84; y2 := TRUE; y3 := FALSE; t0_start := TRUE; t0_up := FALSE;t1_start := FALSE; 
    ELSIF ((x2 = TRUE) AND  ( TRUE ) AND  (x10 = FALSE) AND  (t0.Q = TRUE) AND  ( TRUE )) THEN 
        cstate64 := 87; y2 := TRUE; y3 := TRUE; t0_start := TRUE; t0_up := FALSE;t1_start := TRUE; t1_up := FALSE; 
    ELSIF ((x2 = TRUE) AND  ( TRUE ) AND  (x10 = TRUE) AND  (t0.Q = FALSE) AND  ( TRUE )) THEN 
        cstate64 := 68; y2 := FALSE; y3 := FALSE; t0_start := FALSE;t1_start := FALSE; 
    ELSIF ((x2 = TRUE) AND  ( TRUE ) AND  (x10 = TRUE) AND  (t0.Q = TRUE) AND  ( TRUE )) THEN 
        cstate64 := 65; y2 := FALSE; y3 := FALSE; t0_start := FALSE;t1_start := FALSE; 
    END_IF;
33:
    IF ((x2 = FALSE) AND  ( TRUE ) AND  (x10 = FALSE) AND  (t0.Q = FALSE) AND  (t1.Q = FALSE)) OR ((x2 = FALSE) AND  ( TRUE ) AND  (x10 = TRUE) AND  (t0.Q = FALSE) AND  ( TRUE )) THEN 
        cstate64 := 36; y2 := FALSE; y3 := FALSE; t0_start := FALSE;t1_start := FALSE; 
    ELSIF ((x2 = FALSE) AND  ( TRUE ) AND  (x10 = FALSE) AND  (t0.Q = FALSE) AND  (t1.Q = TRUE)) THEN 
        cstate64 := 36; y2 := FALSE; y3 := FALSE; t0_start := FALSE;t1_start := FALSE; 
    ELSIF ((x2 = FALSE) AND  ( TRUE ) AND  (x10 = FALSE) AND  (t0.Q = TRUE) AND  ( TRUE )) THEN 
        cstate64 := 33; y2 := FALSE; y3 := FALSE; t0_start := FALSE;t1_start := FALSE; 
    ELSIF ((x2 = FALSE) AND  ( TRUE ) AND  (x10 = TRUE) AND  (t0.Q = TRUE) AND  ( TRUE )) THEN 
        cstate64 := 33; y2 := FALSE; y3 := FALSE; t0_start := FALSE;t1_start := FALSE; 
    ELSIF ((x2 = TRUE) AND  ( TRUE ) AND  (x10 = FALSE) AND  (t0.Q = FALSE) AND  (t1.Q = FALSE)) THEN 
        cstate64 := 84; y2 := TRUE; y3 := FALSE; t0_start := TRUE; t0_up := FALSE;t1_start := FALSE; 
    ELSIF ((x2 = TRUE) AND  ( TRUE ) AND  (x10 = FALSE) AND  (t0.Q = FALSE) AND  (t1.Q = TRUE)) THEN 
        cstate64 := 84; y2 := TRUE; y3 := FALSE; t0_start := TRUE; t0_up := FALSE;t1_start := FALSE; 
    ELSIF ((x2 = TRUE) AND  ( TRUE ) AND  (x10 = FALSE) AND  (t0.Q = TRUE) AND  ( TRUE )) THEN 
        cstate64 := 81; y2 := TRUE; y3 := FALSE; t0_start := TRUE; t0_up := FALSE;t1_start := FALSE; 
    ELSIF ((x2 = TRUE) AND  ( TRUE ) AND  (x10 = TRUE) AND  (t0.Q = FALSE) AND  ( TRUE )) THEN 
        cstate64 := 68; y2 := FALSE; y3 := FALSE; t0_start := FALSE;t1_start := FALSE; 
    ELSIF ((x2 = TRUE) AND  ( TRUE ) AND  (x10 = TRUE) AND  (t0.Q = TRUE) AND  ( TRUE )) THEN 
        cstate64 := 65; y2 := FALSE; y3 := FALSE; t0_start := FALSE;t1_start := FALSE; 
    END_IF;
34:
    IF ((x2 = FALSE) AND  ( TRUE ) AND  ( TRUE ) AND  (t0.Q = FALSE) AND  (t1.Q = FALSE)) THEN 
        cstate64 := 35; y2 := FALSE; y3 := FALSE; t0_start := FALSE;t1_start := FALSE; 
    ELSIF ((x2 = FALSE) AND  ( TRUE ) AND  (x10 = FALSE) AND  (t0.Q = FALSE) AND  (t1.Q = TRUE)) THEN 
        cstate64 := 36; y2 := FALSE; y3 := FALSE; t0_start := FALSE;t1_start := FALSE; 
    ELSIF ((x2 = FALSE) AND  ( TRUE ) AND  (x10 = FALSE) AND  (t0.Q = TRUE) AND  (t1.Q = FALSE)) THEN 
        cstate64 := 34; y2 := FALSE; y3 := FALSE; t0_start := FALSE;t1_start := FALSE; 
    ELSIF ((x2 = FALSE) AND  ( TRUE ) AND  (x10 = FALSE) AND  (t0.Q = TRUE) AND  (t1.Q = TRUE)) THEN 
        cstate64 := 33; y2 := FALSE; y3 := FALSE; t0_start := FALSE;t1_start := FALSE; 
    ELSIF ((x2 = FALSE) AND  ( TRUE ) AND  (x10 = TRUE) AND  (t0.Q = FALSE) AND  (t1.Q = TRUE)) THEN 
        cstate64 := 36; y2 := FALSE; y3 := FALSE; t0_start := FALSE;t1_start := FALSE; 
    ELSIF ((x2 = FALSE) AND  ( TRUE ) AND  (x10 = TRUE) AND  (t0.Q = TRUE) AND  (t1.Q = FALSE)) THEN 
        cstate64 := 34; y2 := FALSE; y3 := FALSE; t0_start := FALSE;t1_start := FALSE; 
    ELSIF ((x2 = FALSE) AND  ( TRUE ) AND  (x10 = TRUE) AND  (t0.Q = TRUE) AND  (t1.Q = TRUE)) THEN 
        cstate64 := 33; y2 := FALSE; y3 := FALSE; t0_start := FALSE;t1_start := FALSE; 
    ELSIF ((x2 = TRUE) AND  ( TRUE ) AND  (x10 = FALSE) AND  (t0.Q = FALSE) AND  (t1.Q = FALSE)) THEN 
        cstate64 := 83; y2 := TRUE; y3 := FALSE; t0_start := TRUE; t0_up := FALSE;t1_start := FALSE; 
    ELSIF ((x2 = TRUE) AND  ( TRUE ) AND  (x10 = FALSE) AND  (t0.Q = FALSE) AND  (t1.Q = TRUE)) THEN 
        cstate64 := 84; y2 := TRUE; y3 := FALSE; t0_start := TRUE; t0_up := FALSE;t1_start := FALSE; 
    ELSIF ((x2 = TRUE) AND  ( TRUE ) AND  (x10 = FALSE) AND  (t0.Q = TRUE) AND  (t1.Q = FALSE)) THEN 
        cstate64 := 82; y2 := TRUE; y3 := FALSE; t0_start := TRUE; t0_up := FALSE;t1_start := FALSE; 
    ELSIF ((x2 = TRUE) AND  ( TRUE ) AND  (x10 = FALSE) AND  (t0.Q = TRUE) AND  (t1.Q = TRUE)) THEN 
        cstate64 := 81; y2 := TRUE; y3 := FALSE; t0_start := TRUE; t0_up := FALSE;t1_start := FALSE; 
    ELSIF ((x2 = TRUE) AND  ( TRUE ) AND  (x10 = TRUE) AND  (t0.Q = FALSE) AND  (t1.Q = FALSE)) THEN 
        cstate64 := 67; y2 := FALSE; y3 := FALSE; t0_start := FALSE;t1_start := FALSE; 
    ELSIF ((x2 = TRUE) AND  ( TRUE ) AND  (x10 = TRUE) AND  (t0.Q = FALSE) AND  (t1.Q = TRUE)) THEN 
        cstate64 := 68; y2 := FALSE; y3 := FALSE; t0_start := FALSE;t1_start := FALSE; 
    ELSIF ((x2 = TRUE) AND  ( TRUE ) AND  (x10 = TRUE) AND  (t0.Q = TRUE) AND  (t1.Q = FALSE)) THEN 
        cstate64 := 66; y2 := FALSE; y3 := FALSE; t0_start := FALSE;t1_start := FALSE; 
    ELSIF ((x2 = TRUE) AND  ( TRUE ) AND  (x10 = TRUE) AND  (t0.Q = TRUE) AND  (t1.Q = TRUE)) THEN 
        cstate64 := 65; y2 := FALSE; y3 := FALSE; t0_start := FALSE;t1_start := FALSE; 
    END_IF;
37:
    IF ((x2 = FALSE) AND  ( TRUE ) AND  (x10 = FALSE) AND  (t0.Q = FALSE) AND  (t1.Q = FALSE)) THEN 
        cstate64 := 41; y2 := FALSE; y3 := TRUE; t0_start := FALSE;t1_start := FALSE; 
    ELSIF ((x2 = FALSE) AND  ( TRUE ) AND  (x10 = FALSE) AND  (t0.Q = FALSE) AND  (t1.Q = TRUE)) THEN 
        cstate64 := 36; y2 := FALSE; y3 := FALSE; t0_start := FALSE;t1_start := FALSE; 
    ELSIF ((x2 = FALSE) AND  ( TRUE ) AND  (x10 = FALSE) AND  (t0.Q = TRUE) AND  (t1.Q = FALSE)) THEN 
        cstate64 := 37; y2 := FALSE; y3 := TRUE; t0_start := FALSE;t1_start := FALSE; 
    ELSIF ((x2 = FALSE) AND  ( TRUE ) AND  (x10 = FALSE) AND  (t0.Q = TRUE) AND  (t1.Q = TRUE)) THEN 
        cstate64 := 33; y2 := FALSE; y3 := FALSE; t0_start := FALSE;t1_start := FALSE; 
    ELSIF ((x2 = FALSE) AND  ( TRUE ) AND  (x10 = TRUE) AND  (t0.Q = FALSE) AND  (t1.Q = FALSE)) THEN 
        cstate64 := 35; y2 := FALSE; y3 := FALSE; t0_start := FALSE;t1_start := FALSE; 
    ELSIF ((x2 = FALSE) AND  ( TRUE ) AND  (x10 = TRUE) AND  (t0.Q = FALSE) AND  (t1.Q = TRUE)) THEN 
        cstate64 := 36; y2 := FALSE; y3 := FALSE; t0_start := FALSE;t1_start := FALSE; 
    ELSIF ((x2 = FALSE) AND  ( TRUE ) AND  (x10 = TRUE) AND  (t0.Q = TRUE) AND  (t1.Q = FALSE)) THEN 
        cstate64 := 34; y2 := FALSE; y3 := FALSE; t0_start := FALSE;t1_start := FALSE; 
    ELSIF ((x2 = FALSE) AND  ( TRUE ) AND  (x10 = TRUE) AND  (t0.Q = TRUE) AND  (t1.Q = TRUE)) THEN 
        cstate64 := 33; y2 := FALSE; y3 := FALSE; t0_start := FALSE;t1_start := FALSE; 
    ELSIF ((x2 = TRUE) AND  ( TRUE ) AND  (x10 = FALSE) AND  (t0.Q = FALSE) AND  (t1.Q = FALSE)) THEN 
        cstate64 := 90; y2 := TRUE; y3 := TRUE; t0_start := TRUE; t0_up := FALSE;t1_start := FALSE; 
    ELSIF ((x2 = TRUE) AND  ( TRUE ) AND  (x10 = FALSE) AND  (t0.Q = FALSE) AND  (t1.Q = TRUE)) THEN 
        cstate64 := 84; y2 := TRUE; y3 := FALSE; t0_start := TRUE; t0_up := FALSE;t1_start := FALSE; 
    ELSIF ((x2 = TRUE) AND  ( TRUE ) AND  (x10 = FALSE) AND  (t0.Q = TRUE) AND  (t1.Q = FALSE)) THEN 
        cstate64 := 86; y2 := TRUE; y3 := TRUE; t0_start := TRUE; t0_up := FALSE;t1_start := FALSE; 
    ELSIF ((x2 = TRUE) AND  ( TRUE ) AND  (x10 = FALSE) AND  (t0.Q = TRUE) AND  (t1.Q = TRUE)) THEN 
        cstate64 := 81; y2 := TRUE; y3 := FALSE; t0_start := TRUE; t0_up := FALSE;t1_start := FALSE; 
    ELSIF ((x2 = TRUE) AND  ( TRUE ) AND  (x10 = TRUE) AND  (t0.Q = FALSE) AND  (t1.Q = FALSE)) THEN 
        cstate64 := 67; y2 := FALSE; y3 := FALSE; t0_start := FALSE;t1_start := FALSE; 
    ELSIF ((x2 = TRUE) AND  ( TRUE ) AND  (x10 = TRUE) AND  (t0.Q = FALSE) AND  (t1.Q = TRUE)) THEN 
        cstate64 := 68; y2 := FALSE; y3 := FALSE; t0_start := FALSE;t1_start := FALSE; 
    ELSIF ((x2 = TRUE) AND  ( TRUE ) AND  (x10 = TRUE) AND  (t0.Q = TRUE) AND  (t1.Q = FALSE)) THEN 
        cstate64 := 66; y2 := FALSE; y3 := FALSE; t0_start := FALSE;t1_start := FALSE; 
    ELSIF ((x2 = TRUE) AND  ( TRUE ) AND  (x10 = TRUE) AND  (t0.Q = TRUE) AND  (t1.Q = TRUE)) THEN 
        cstate64 := 65; y2 := FALSE; y3 := FALSE; t0_start := FALSE;t1_start := FALSE; 
    END_IF;
20:
    IF ((x2 = FALSE) AND  ( TRUE ) AND  (x10 = FALSE) AND  (t0.Q = FALSE) AND  (t1.Q = FALSE)) OR ((x2 = FALSE) AND  ( TRUE ) AND  (x10 = TRUE) AND  (t0.Q = FALSE) AND  ( TRUE )) THEN 
        cstate64 := 20; y2 := FALSE; y3 := FALSE; t0_start := FALSE;t1_start := FALSE; 
    ELSIF ((x2 = FALSE) AND  ( TRUE ) AND  (x10 = FALSE) AND  (t0.Q = FALSE) AND  (t1.Q = TRUE)) THEN 
        cstate64 := 20; y2 := FALSE; y3 := FALSE; t0_start := FALSE;t1_start := FALSE; 
    ELSIF ((x2 = FALSE) AND  ( TRUE ) AND  (x10 = FALSE) AND  (t0.Q = TRUE) AND  ( TRUE )) THEN 
        cstate64 := 40; y2 := FALSE; y3 := TRUE; t0_start := FALSE;t1_start := TRUE; t1_up := FALSE; 
    ELSIF ((x2 = FALSE) AND  ( TRUE ) AND  (x10 = TRUE) AND  (t0.Q = TRUE) AND  ( TRUE )) THEN 
        cstate64 := 33; y2 := FALSE; y3 := FALSE; t0_start := FALSE;t1_start := FALSE; 
    ELSIF ((x2 = TRUE) AND  ( TRUE ) AND  (x10 = FALSE) AND  (t0.Q = FALSE) AND  (t1.Q = FALSE)) THEN 
        cstate64 := 84; y2 := TRUE; y3 := FALSE; t0_start := TRUE; t0_up := FALSE;t1_start := FALSE; 
    ELSIF ((x2 = TRUE) AND  ( TRUE ) AND  (x10 = FALSE) AND  (t0.Q = FALSE) AND  (t1.Q = TRUE)) THEN 
        cstate64 := 84; y2 := TRUE; y3 := FALSE; t0_start := TRUE; t0_up := FALSE;t1_start := FALSE; 
    ELSIF ((x2 = TRUE) AND  ( TRUE ) AND  (x10 = FALSE) AND  (t0.Q = TRUE) AND  ( TRUE )) THEN 
        cstate64 := 87; y2 := TRUE; y3 := TRUE; t0_start := TRUE; t0_up := FALSE;t1_start := TRUE; t1_up := FALSE; 
    ELSIF ((x2 = TRUE) AND  ( TRUE ) AND  (x10 = TRUE) AND  (t0.Q = FALSE) AND  ( TRUE )) THEN 
        cstate64 := 52; y2 := FALSE; y3 := FALSE; t0_start := FALSE;t1_start := FALSE; 
    ELSIF ((x2 = TRUE) AND  ( TRUE ) AND  (x10 = TRUE) AND  (t0.Q = TRUE) AND  ( TRUE )) THEN 
        cstate64 := 65; y2 := FALSE; y3 := FALSE; t0_start := FALSE;t1_start := FALSE; 
    END_IF;
41:
    IF ((x2 = FALSE) AND  ( TRUE ) AND  (x10 = FALSE) AND  (t0.Q = FALSE) AND  (t1.Q = FALSE)) THEN 
        cstate64 := 41; y2 := FALSE; y3 := TRUE; t0_start := FALSE;t1_start := FALSE; 
    ELSIF ((x2 = FALSE) AND  ( TRUE ) AND  (x10 = FALSE) AND  (t0.Q = FALSE) AND  (t1.Q = TRUE)) THEN 
        cstate64 := 36; y2 := FALSE; y3 := FALSE; t0_start := FALSE;t1_start := FALSE; 
    ELSIF ((x2 = FALSE) AND  ( TRUE ) AND  (x10 = FALSE) AND  (t0.Q = TRUE) AND  ( TRUE )) THEN 
        cstate64 := 37; y2 := FALSE; y3 := TRUE; t0_start := FALSE;t1_start := TRUE; t1_up := FALSE; 
    ELSIF ((x2 = FALSE) AND  ( TRUE ) AND  (x10 = TRUE) AND  (t0.Q = FALSE) AND  (t1.Q = FALSE)) THEN 
        cstate64 := 35; y2 := FALSE; y3 := FALSE; t0_start := FALSE;t1_start := FALSE; 
    ELSIF ((x2 = FALSE) AND  ( TRUE ) AND  (x10 = TRUE) AND  (t0.Q = FALSE) AND  (t1.Q = TRUE)) THEN 
        cstate64 := 36; y2 := FALSE; y3 := FALSE; t0_start := FALSE;t1_start := FALSE; 
    ELSIF ((x2 = FALSE) AND  ( TRUE ) AND  (x10 = TRUE) AND  (t0.Q = TRUE) AND  (t1.Q = FALSE)) THEN 
        cstate64 := 34; y2 := FALSE; y3 := FALSE; t0_start := FALSE;t1_start := FALSE; 
    ELSIF ((x2 = FALSE) AND  ( TRUE ) AND  (x10 = TRUE) AND  (t0.Q = TRUE) AND  (t1.Q = TRUE)) THEN 
        cstate64 := 33; y2 := FALSE; y3 := FALSE; t0_start := FALSE;t1_start := FALSE; 
    ELSIF ((x2 = TRUE) AND  ( TRUE ) AND  (x10 = FALSE) AND  (t0.Q = FALSE) AND  (t1.Q = FALSE)) THEN 
        cstate64 := 90; y2 := TRUE; y3 := TRUE; t0_start := TRUE; t0_up := FALSE;t1_start := FALSE; 
    ELSIF ((x2 = TRUE) AND  ( TRUE ) AND  (x10 = FALSE) AND  (t0.Q = FALSE) AND  (t1.Q = TRUE)) THEN 
        cstate64 := 84; y2 := TRUE; y3 := FALSE; t0_start := TRUE; t0_up := FALSE;t1_start := FALSE; 
    ELSIF ((x2 = TRUE) AND  ( TRUE ) AND  (x10 = FALSE) AND  (t0.Q = TRUE) AND  ( TRUE )) THEN 
        cstate64 := 86; y2 := TRUE; y3 := TRUE; t0_start := TRUE; t0_up := FALSE;t1_start := TRUE; t1_up := FALSE; 
    ELSIF ((x2 = TRUE) AND  ( TRUE ) AND  (x10 = TRUE) AND  (t0.Q = FALSE) AND  (t1.Q = FALSE)) THEN 
        cstate64 := 67; y2 := FALSE; y3 := FALSE; t0_start := FALSE;t1_start := FALSE; 
    ELSIF ((x2 = TRUE) AND  ( TRUE ) AND  (x10 = TRUE) AND  (t0.Q = FALSE) AND  (t1.Q = TRUE)) THEN 
        cstate64 := 68; y2 := FALSE; y3 := FALSE; t0_start := FALSE;t1_start := FALSE; 
    ELSIF ((x2 = TRUE) AND  ( TRUE ) AND  (x10 = TRUE) AND  (t0.Q = TRUE) AND  (t1.Q = FALSE)) THEN 
        cstate64 := 66; y2 := FALSE; y3 := FALSE; t0_start := FALSE;t1_start := FALSE; 
    ELSIF ((x2 = TRUE) AND  ( TRUE ) AND  (x10 = TRUE) AND  (t0.Q = TRUE) AND  (t1.Q = TRUE)) THEN 
        cstate64 := 65; y2 := FALSE; y3 := FALSE; t0_start := FALSE;t1_start := FALSE; 
    END_IF;
107:
    IF ((x2 = FALSE) AND  ( TRUE ) AND  (x10 = FALSE) AND  (t0.Q = FALSE) AND  (t1.Q = FALSE)) THEN 
        cstate64 := 107; y2 := TRUE; y3 := TRUE; t0_start := FALSE;t1_start := FALSE; 
    ELSIF ((x2 = FALSE) AND  ( TRUE ) AND  (x10 = FALSE) AND  (t0.Q = FALSE) AND  (t1.Q = TRUE)) THEN 
        cstate64 := 100; y2 := TRUE; y3 := FALSE; t0_start := FALSE;t1_start := FALSE; 
    ELSIF ((x2 = FALSE) AND  ( TRUE ) AND  (x10 = FALSE) AND  (t0.Q = TRUE) AND  (t1.Q = FALSE)) THEN 
        cstate64 := 40; y2 := FALSE; y3 := TRUE; t0_start := FALSE;t1_start := TRUE; t1_up := FALSE; 
    ELSIF ((x2 = FALSE) AND  ( TRUE ) AND  (x10 = FALSE) AND  (t0.Q = TRUE) AND  (t1.Q = TRUE)) THEN 
        cstate64 := 37; y2 := FALSE; y3 := TRUE; t0_start := FALSE;t1_start := TRUE; t1_up := FALSE; 
    ELSIF ((x2 = FALSE) AND  ( TRUE ) AND  (x10 = TRUE) AND  (t0.Q = FALSE) AND  (t1.Q = FALSE)) THEN 
        cstate64 := 19; y2 := FALSE; y3 := FALSE; t0_start := FALSE;t1_start := FALSE; 
    ELSIF ((x2 = FALSE) AND  ( TRUE ) AND  (x10 = TRUE) AND  (t0.Q = FALSE) AND  (t1.Q = TRUE)) THEN 
        cstate64 := 20; y2 := FALSE; y3 := FALSE; t0_start := FALSE;t1_start := FALSE; 
    ELSIF ((x2 = FALSE) AND  ( TRUE ) AND  (x10 = TRUE) AND  (t0.Q = TRUE) AND  (t1.Q = FALSE)) THEN 
        cstate64 := 34; y2 := FALSE; y3 := FALSE; t0_start := FALSE;t1_start := FALSE; 
    ELSIF ((x2 = FALSE) AND  ( TRUE ) AND  (x10 = TRUE) AND  (t0.Q = TRUE) AND  (t1.Q = TRUE)) THEN 
        cstate64 := 33; y2 := FALSE; y3 := FALSE; t0_start := FALSE;t1_start := FALSE; 
    ELSIF ((x2 = TRUE) AND  ( TRUE ) AND  (x10 = FALSE) AND  (t0.Q = FALSE) AND  (t1.Q = FALSE)) THEN 
        cstate64 := 91; y2 := TRUE; y3 := TRUE; t0_start := TRUE; t0_up := FALSE;t1_start := FALSE; 
    ELSIF ((x2 = TRUE) AND  ( TRUE ) AND  (x10 = FALSE) AND  (t0.Q = FALSE) AND  (t1.Q = TRUE)) THEN 
        cstate64 := 84; y2 := TRUE; y3 := FALSE; t0_start := TRUE; t0_up := FALSE;t1_start := FALSE; 
    ELSIF ((x2 = TRUE) AND  ( TRUE ) AND  (x10 = FALSE) AND  (t0.Q = TRUE) AND  (t1.Q = FALSE)) THEN 
        cstate64 := 87; y2 := TRUE; y3 := TRUE; t0_start := TRUE; t0_up := FALSE;t1_start := TRUE; t1_up := FALSE; 
    ELSIF ((x2 = TRUE) AND  ( TRUE ) AND  (x10 = FALSE) AND  (t0.Q = TRUE) AND  (t1.Q = TRUE)) THEN 
        cstate64 := 86; y2 := TRUE; y3 := TRUE; t0_start := TRUE; t0_up := FALSE;t1_start := TRUE; t1_up := FALSE; 
    ELSIF ((x2 = TRUE) AND  ( TRUE ) AND  (x10 = TRUE) AND  (t0.Q = FALSE) AND  (t1.Q = FALSE)) THEN 
        cstate64 := 51; y2 := FALSE; y3 := FALSE; t0_start := FALSE;t1_start := FALSE; 
    ELSIF ((x2 = TRUE) AND  ( TRUE ) AND  (x10 = TRUE) AND  (t0.Q = FALSE) AND  (t1.Q = TRUE)) THEN 
        cstate64 := 52; y2 := FALSE; y3 := FALSE; t0_start := FALSE;t1_start := FALSE; 
    ELSIF ((x2 = TRUE) AND  ( TRUE ) AND  (x10 = TRUE) AND  (t0.Q = TRUE) AND  (t1.Q = FALSE)) THEN 
        cstate64 := 66; y2 := FALSE; y3 := FALSE; t0_start := FALSE;t1_start := FALSE; 
    ELSIF ((x2 = TRUE) AND  ( TRUE ) AND  (x10 = TRUE) AND  (t0.Q = TRUE) AND  (t1.Q = TRUE)) THEN 
        cstate64 := 65; y2 := FALSE; y3 := FALSE; t0_start := FALSE;t1_start := FALSE; 
    END_IF;
40:
    IF ((x2 = FALSE) AND  ( TRUE ) AND  (x10 = FALSE) AND  (t0.Q = FALSE) AND  (t1.Q = FALSE)) THEN 
        cstate64 := 44; y2 := FALSE; y3 := TRUE; t0_start := FALSE;t1_start := FALSE; 
    ELSIF ((x2 = FALSE) AND  ( TRUE ) AND  (x10 = FALSE) AND  (t0.Q = FALSE) AND  (t1.Q = TRUE)) THEN 
        cstate64 := 36; y2 := FALSE; y3 := FALSE; t0_start := FALSE;t1_start := FALSE; 
    ELSIF ((x2 = FALSE) AND  ( TRUE ) AND  (x10 = FALSE) AND  (t0.Q = TRUE) AND  (t1.Q = FALSE)) THEN 
        cstate64 := 40; y2 := FALSE; y3 := TRUE; t0_start := FALSE;t1_start := FALSE; 
    ELSIF ((x2 = FALSE) AND  ( TRUE ) AND  (x10 = FALSE) AND  (t0.Q = TRUE) AND  (t1.Q = TRUE)) THEN 
        cstate64 := 33; y2 := FALSE; y3 := FALSE; t0_start := FALSE;t1_start := FALSE; 
    ELSIF ((x2 = FALSE) AND  ( TRUE ) AND  (x10 = TRUE) AND  (t0.Q = FALSE) AND  (t1.Q = FALSE)) THEN 
        cstate64 := 35; y2 := FALSE; y3 := FALSE; t0_start := FALSE;t1_start := FALSE; 
    ELSIF ((x2 = FALSE) AND  ( TRUE ) AND  (x10 = TRUE) AND  (t0.Q = FALSE) AND  (t1.Q = TRUE)) THEN 
        cstate64 := 36; y2 := FALSE; y3 := FALSE; t0_start := FALSE;t1_start := FALSE; 
    ELSIF ((x2 = FALSE) AND  ( TRUE ) AND  (x10 = TRUE) AND  (t0.Q = TRUE) AND  (t1.Q = FALSE)) THEN 
        cstate64 := 34; y2 := FALSE; y3 := FALSE; t0_start := FALSE;t1_start := FALSE; 
    ELSIF ((x2 = FALSE) AND  ( TRUE ) AND  (x10 = TRUE) AND  (t0.Q = TRUE) AND  (t1.Q = TRUE)) THEN 
        cstate64 := 33; y2 := FALSE; y3 := FALSE; t0_start := FALSE;t1_start := FALSE; 
    ELSIF ((x2 = TRUE) AND  ( TRUE ) AND  (x10 = FALSE) AND  (t0.Q = FALSE) AND  (t1.Q = FALSE)) THEN 
        cstate64 := 91; y2 := TRUE; y3 := TRUE; t0_start := TRUE; t0_up := FALSE;t1_start := FALSE; 
    ELSIF ((x2 = TRUE) AND  ( TRUE ) AND  (x10 = FALSE) AND  (t0.Q = FALSE) AND  (t1.Q = TRUE)) THEN 
        cstate64 := 84; y2 := TRUE; y3 := FALSE; t0_start := TRUE; t0_up := FALSE;t1_start := FALSE; 
    ELSIF ((x2 = TRUE) AND  ( TRUE ) AND  (x10 = FALSE) AND  (t0.Q = TRUE) AND  (t1.Q = FALSE)) THEN 
        cstate64 := 87; y2 := TRUE; y3 := TRUE; t0_start := TRUE; t0_up := FALSE;t1_start := FALSE; 
    ELSIF ((x2 = TRUE) AND  ( TRUE ) AND  (x10 = FALSE) AND  (t0.Q = TRUE) AND  (t1.Q = TRUE)) THEN 
        cstate64 := 81; y2 := TRUE; y3 := FALSE; t0_start := TRUE; t0_up := FALSE;t1_start := FALSE; 
    ELSIF ((x2 = TRUE) AND  ( TRUE ) AND  (x10 = TRUE) AND  (t0.Q = FALSE) AND  (t1.Q = FALSE)) THEN 
        cstate64 := 67; y2 := FALSE; y3 := FALSE; t0_start := FALSE;t1_start := FALSE; 
    ELSIF ((x2 = TRUE) AND  ( TRUE ) AND  (x10 = TRUE) AND  (t0.Q = FALSE) AND  (t1.Q = TRUE)) THEN 
        cstate64 := 68; y2 := FALSE; y3 := FALSE; t0_start := FALSE;t1_start := FALSE; 
    ELSIF ((x2 = TRUE) AND  ( TRUE ) AND  (x10 = TRUE) AND  (t0.Q = TRUE) AND  (t1.Q = FALSE)) THEN 
        cstate64 := 66; y2 := FALSE; y3 := FALSE; t0_start := FALSE;t1_start := FALSE; 
    ELSIF ((x2 = TRUE) AND  ( TRUE ) AND  (x10 = TRUE) AND  (t0.Q = TRUE) AND  (t1.Q = TRUE)) THEN 
        cstate64 := 65; y2 := FALSE; y3 := FALSE; t0_start := FALSE;t1_start := FALSE; 
    END_IF;
106:
    IF ((x2 = FALSE) AND  ( TRUE ) AND  (x10 = FALSE) AND  (t0.Q = FALSE) AND  (t1.Q = FALSE)) THEN 
        cstate64 := 106; y2 := TRUE; y3 := TRUE; t0_start := FALSE;t1_start := FALSE; 
    ELSIF ((x2 = FALSE) AND  ( TRUE ) AND  (x10 = FALSE) AND  (t0.Q = FALSE) AND  (t1.Q = TRUE)) THEN 
        cstate64 := 100; y2 := TRUE; y3 := FALSE; t0_start := FALSE;t1_start := FALSE; 
    ELSIF ((x2 = FALSE) AND  ( TRUE ) AND  (x10 = FALSE) AND  (t0.Q = TRUE) AND  ( TRUE )) THEN 
        cstate64 := 37; y2 := FALSE; y3 := TRUE; t0_start := FALSE;t1_start := TRUE; t1_up := FALSE; 
    ELSIF ((x2 = FALSE) AND  ( TRUE ) AND  (x10 = TRUE) AND  (t0.Q = FALSE) AND  (t1.Q = FALSE)) THEN 
        cstate64 := 19; y2 := FALSE; y3 := FALSE; t0_start := FALSE;t1_start := FALSE; 
    ELSIF ((x2 = FALSE) AND  ( TRUE ) AND  (x10 = TRUE) AND  (t0.Q = FALSE) AND  (t1.Q = TRUE)) THEN 
        cstate64 := 20; y2 := FALSE; y3 := FALSE; t0_start := FALSE;t1_start := FALSE; 
    ELSIF ((x2 = FALSE) AND  ( TRUE ) AND  (x10 = TRUE) AND  (t0.Q = TRUE) AND  (t1.Q = FALSE)) THEN 
        cstate64 := 34; y2 := FALSE; y3 := FALSE; t0_start := FALSE;t1_start := FALSE; 
    ELSIF ((x2 = FALSE) AND  ( TRUE ) AND  (x10 = TRUE) AND  (t0.Q = TRUE) AND  (t1.Q = TRUE)) THEN 
        cstate64 := 33; y2 := FALSE; y3 := FALSE; t0_start := FALSE;t1_start := FALSE; 
    ELSIF ((x2 = TRUE) AND  ( TRUE ) AND  (x10 = FALSE) AND  (t0.Q = FALSE) AND  (t1.Q = FALSE)) THEN 
        cstate64 := 90; y2 := TRUE; y3 := TRUE; t0_start := TRUE; t0_up := FALSE;t1_start := FALSE; 
    ELSIF ((x2 = TRUE) AND  ( TRUE ) AND  (x10 = FALSE) AND  (t0.Q = FALSE) AND  (t1.Q = TRUE)) THEN 
        cstate64 := 84; y2 := TRUE; y3 := FALSE; t0_start := TRUE; t0_up := FALSE;t1_start := FALSE; 
    ELSIF ((x2 = TRUE) AND  ( TRUE ) AND  (x10 = FALSE) AND  (t0.Q = TRUE) AND  ( TRUE )) THEN 
        cstate64 := 86; y2 := TRUE; y3 := TRUE; t0_start := TRUE; t0_up := FALSE;t1_start := TRUE; t1_up := FALSE; 
    ELSIF ((x2 = TRUE) AND  ( TRUE ) AND  (x10 = TRUE) AND  (t0.Q = FALSE) AND  (t1.Q = FALSE)) THEN 
        cstate64 := 51; y2 := FALSE; y3 := FALSE; t0_start := FALSE;t1_start := FALSE; 
    ELSIF ((x2 = TRUE) AND  ( TRUE ) AND  (x10 = TRUE) AND  (t0.Q = FALSE) AND  (t1.Q = TRUE)) THEN 
        cstate64 := 52; y2 := FALSE; y3 := FALSE; t0_start := FALSE;t1_start := FALSE; 
    ELSIF ((x2 = TRUE) AND  ( TRUE ) AND  (x10 = TRUE) AND  (t0.Q = TRUE) AND  (t1.Q = FALSE)) THEN 
        cstate64 := 66; y2 := FALSE; y3 := FALSE; t0_start := FALSE;t1_start := FALSE; 
    ELSIF ((x2 = TRUE) AND  ( TRUE ) AND  (x10 = TRUE) AND  (t0.Q = TRUE) AND  (t1.Q = TRUE)) THEN 
        cstate64 := 65; y2 := FALSE; y3 := FALSE; t0_start := FALSE;t1_start := FALSE; 
    END_IF;
82:
    IF ((x2 = FALSE) AND  ( TRUE ) AND  (x10 = FALSE) AND  (t0.Q = FALSE) AND  (t1.Q = FALSE)) THEN 
        cstate64 := 99; y2 := TRUE; y3 := FALSE; t0_start := FALSE;t1_start := FALSE; 
    ELSIF ((x2 = FALSE) AND  ( TRUE ) AND  (x10 = FALSE) AND  (t0.Q = FALSE) AND  (t1.Q = TRUE)) THEN 
        cstate64 := 100; y2 := TRUE; y3 := FALSE; t0_start := FALSE;t1_start := FALSE; 
    ELSIF ((x2 = FALSE) AND  ( TRUE ) AND  (x10 = FALSE) AND  (t0.Q = TRUE) AND  (t1.Q = FALSE)) THEN 
        cstate64 := 34; y2 := FALSE; y3 := FALSE; t0_start := FALSE;t1_start := FALSE; 
    ELSIF ((x2 = FALSE) AND  ( TRUE ) AND  (x10 = FALSE) AND  (t0.Q = TRUE) AND  (t1.Q = TRUE)) THEN 
        cstate64 := 33; y2 := FALSE; y3 := FALSE; t0_start := FALSE;t1_start := FALSE; 
    ELSIF ((x2 = FALSE) AND  ( TRUE ) AND  (x10 = TRUE) AND  (t0.Q = FALSE) AND  (t1.Q = FALSE)) THEN 
        cstate64 := 19; y2 := FALSE; y3 := FALSE; t0_start := FALSE;t1_start := FALSE; 
    ELSIF ((x2 = FALSE) AND  ( TRUE ) AND  (x10 = TRUE) AND  (t0.Q = FALSE) AND  (t1.Q = TRUE)) THEN 
        cstate64 := 20; y2 := FALSE; y3 := FALSE; t0_start := FALSE;t1_start := FALSE; 
    ELSIF ((x2 = FALSE) AND  ( TRUE ) AND  (x10 = TRUE) AND  (t0.Q = TRUE) AND  (t1.Q = FALSE)) THEN 
        cstate64 := 34; y2 := FALSE; y3 := FALSE; t0_start := FALSE;t1_start := FALSE; 
    ELSIF ((x2 = FALSE) AND  ( TRUE ) AND  (x10 = TRUE) AND  (t0.Q = TRUE) AND  (t1.Q = TRUE)) THEN 
        cstate64 := 33; y2 := FALSE; y3 := FALSE; t0_start := FALSE;t1_start := FALSE; 
    ELSIF ((x2 = TRUE) AND  ( TRUE ) AND  (x10 = FALSE) AND  (t0.Q = FALSE) AND  (t1.Q = FALSE)) THEN 
        cstate64 := 83; y2 := TRUE; y3 := FALSE; t0_start := FALSE;t1_start := FALSE; 
    ELSIF ((x2 = TRUE) AND  ( TRUE ) AND  (x10 = FALSE) AND  (t0.Q = FALSE) AND  (t1.Q = TRUE)) THEN 
        cstate64 := 84; y2 := TRUE; y3 := FALSE; t0_start := FALSE;t1_start := FALSE; 
    ELSIF ((x2 = TRUE) AND  ( TRUE ) AND  ( TRUE ) AND  (t0.Q = TRUE) AND  (t1.Q = FALSE)) THEN 
        cstate64 := 66; y2 := FALSE; y3 := FALSE; t0_start := FALSE;t1_start := FALSE; 
    ELSIF ((x2 = TRUE) AND  ( TRUE ) AND  ( TRUE ) AND  (t0.Q = TRUE) AND  (t1.Q = TRUE)) THEN 
        cstate64 := 65; y2 := FALSE; y3 := FALSE; t0_start := FALSE;t1_start := FALSE; 
    ELSIF ((x2 = TRUE) AND  ( TRUE ) AND  (x10 = TRUE) AND  (t0.Q = FALSE) AND  (t1.Q = FALSE)) THEN 
        cstate64 := 51; y2 := FALSE; y3 := FALSE; t0_start := FALSE;t1_start := FALSE; 
    ELSIF ((x2 = TRUE) AND  ( TRUE ) AND  (x10 = TRUE) AND  (t0.Q = FALSE) AND  (t1.Q = TRUE)) THEN 
        cstate64 := 52; y2 := FALSE; y3 := FALSE; t0_start := FALSE;t1_start := FALSE; 
    END_IF;
65:
    IF ((x2 = FALSE) AND  ( TRUE ) AND  (x10 = FALSE) AND  (t0.Q = FALSE) AND  (t1.Q = FALSE)) OR ((x2 = FALSE) AND  ( TRUE ) AND  (x10 = TRUE) AND  (t0.Q = FALSE) AND  ( TRUE )) THEN 
        cstate64 := 36; y2 := FALSE; y3 := FALSE; t0_start := FALSE;t1_start := FALSE; 
    ELSIF ((x2 = FALSE) AND  ( TRUE ) AND  (x10 = FALSE) AND  (t0.Q = FALSE) AND  (t1.Q = TRUE)) THEN 
        cstate64 := 36; y2 := FALSE; y3 := FALSE; t0_start := FALSE;t1_start := FALSE; 
    ELSIF ((x2 = FALSE) AND  ( TRUE ) AND  (x10 = FALSE) AND  (t0.Q = TRUE) AND  ( TRUE )) THEN 
        cstate64 := 33; y2 := FALSE; y3 := FALSE; t0_start := FALSE;t1_start := FALSE; 
    ELSIF ((x2 = FALSE) AND  ( TRUE ) AND  (x10 = TRUE) AND  (t0.Q = TRUE) AND  ( TRUE )) THEN 
        cstate64 := 33; y2 := FALSE; y3 := FALSE; t0_start := FALSE;t1_start := FALSE; 
    ELSIF ((x2 = TRUE) AND  ( TRUE ) AND  (x10 = FALSE) AND  (t0.Q = FALSE) AND  (t1.Q = FALSE)) OR ((x2 = TRUE) AND  ( TRUE ) AND  (x10 = TRUE) AND  (t0.Q = FALSE) AND  ( TRUE )) THEN 
        cstate64 := 68; y2 := FALSE; y3 := FALSE; t0_start := FALSE;t1_start := FALSE; 
    ELSIF ((x2 = TRUE) AND  ( TRUE ) AND  (x10 = FALSE) AND  (t0.Q = FALSE) AND  (t1.Q = TRUE)) THEN 
        cstate64 := 68; y2 := FALSE; y3 := FALSE; t0_start := FALSE;t1_start := FALSE; 
    ELSIF ((x2 = TRUE) AND  ( TRUE ) AND  ( TRUE ) AND  (t0.Q = TRUE) AND  ( TRUE )) THEN 
        cstate64 := 65; y2 := FALSE; y3 := FALSE; t0_start := FALSE;t1_start := FALSE; 
    END_IF;
83:
    IF ((x2 = FALSE) AND  ( TRUE ) AND  (x10 = FALSE) AND  (t0.Q = FALSE) AND  (t1.Q = FALSE)) THEN 
        cstate64 := 99; y2 := TRUE; y3 := FALSE; t0_start := FALSE;t1_start := FALSE; 
    ELSIF ((x2 = FALSE) AND  ( TRUE ) AND  (x10 = FALSE) AND  (t0.Q = FALSE) AND  (t1.Q = TRUE)) THEN 
        cstate64 := 100; y2 := TRUE; y3 := FALSE; t0_start := FALSE;t1_start := FALSE; 
    ELSIF ((x2 = FALSE) AND  ( TRUE ) AND  (x10 = FALSE) AND  (t0.Q = TRUE) AND  ( TRUE )) THEN 
        cstate64 := 37; y2 := FALSE; y3 := TRUE; t0_start := FALSE;t1_start := TRUE; t1_up := FALSE; 
    ELSIF ((x2 = FALSE) AND  ( TRUE ) AND  (x10 = TRUE) AND  (t0.Q = FALSE) AND  (t1.Q = FALSE)) THEN 
        cstate64 := 19; y2 := FALSE; y3 := FALSE; t0_start := FALSE;t1_start := FALSE; 
    ELSIF ((x2 = FALSE) AND  ( TRUE ) AND  (x10 = TRUE) AND  (t0.Q = FALSE) AND  (t1.Q = TRUE)) THEN 
        cstate64 := 20; y2 := FALSE; y3 := FALSE; t0_start := FALSE;t1_start := FALSE; 
    ELSIF ((x2 = FALSE) AND  ( TRUE ) AND  (x10 = TRUE) AND  (t0.Q = TRUE) AND  (t1.Q = FALSE)) THEN 
        cstate64 := 34; y2 := FALSE; y3 := FALSE; t0_start := FALSE;t1_start := FALSE; 
    ELSIF ((x2 = FALSE) AND  ( TRUE ) AND  (x10 = TRUE) AND  (t0.Q = TRUE) AND  (t1.Q = TRUE)) THEN 
        cstate64 := 33; y2 := FALSE; y3 := FALSE; t0_start := FALSE;t1_start := FALSE; 
    ELSIF ((x2 = TRUE) AND  ( TRUE ) AND  (x10 = FALSE) AND  (t0.Q = FALSE) AND  (t1.Q = FALSE)) THEN 
        cstate64 := 83; y2 := TRUE; y3 := FALSE; t0_start := FALSE;t1_start := FALSE; 
    ELSIF ((x2 = TRUE) AND  ( TRUE ) AND  (x10 = FALSE) AND  (t0.Q = FALSE) AND  (t1.Q = TRUE)) THEN 
        cstate64 := 84; y2 := TRUE; y3 := FALSE; t0_start := FALSE;t1_start := FALSE; 
    ELSIF ((x2 = TRUE) AND  ( TRUE ) AND  (x10 = FALSE) AND  (t0.Q = TRUE) AND  ( TRUE )) THEN 
        cstate64 := 69; y2 := FALSE; y3 := TRUE; t0_start := FALSE;t1_start := TRUE; t1_up := FALSE; 
    ELSIF ((x2 = TRUE) AND  ( TRUE ) AND  (x10 = TRUE) AND  (t0.Q = FALSE) AND  (t1.Q = FALSE)) THEN 
        cstate64 := 51; y2 := FALSE; y3 := FALSE; t0_start := FALSE;t1_start := FALSE; 
    ELSIF ((x2 = TRUE) AND  ( TRUE ) AND  (x10 = TRUE) AND  (t0.Q = FALSE) AND  (t1.Q = TRUE)) THEN 
        cstate64 := 52; y2 := FALSE; y3 := FALSE; t0_start := FALSE;t1_start := FALSE; 
    ELSIF ((x2 = TRUE) AND  ( TRUE ) AND  (x10 = TRUE) AND  (t0.Q = TRUE) AND  (t1.Q = FALSE)) THEN 
        cstate64 := 66; y2 := FALSE; y3 := FALSE; t0_start := FALSE;t1_start := FALSE; 
    ELSIF ((x2 = TRUE) AND  ( TRUE ) AND  (x10 = TRUE) AND  (t0.Q = TRUE) AND  (t1.Q = TRUE)) THEN 
        cstate64 := 65; y2 := FALSE; y3 := FALSE; t0_start := FALSE;t1_start := FALSE; 
    END_IF;
81:
    IF ((x2 = FALSE) AND  ( TRUE ) AND  (x10 = FALSE) AND  (t0.Q = FALSE) AND  (t1.Q = FALSE)) THEN 
        cstate64 := 100; y2 := TRUE; y3 := FALSE; t0_start := FALSE;t1_start := FALSE; 
    ELSIF ((x2 = FALSE) AND  ( TRUE ) AND  (x10 = FALSE) AND  (t0.Q = FALSE) AND  (t1.Q = TRUE)) THEN 
        cstate64 := 100; y2 := TRUE; y3 := FALSE; t0_start := FALSE;t1_start := FALSE; 
    ELSIF ((x2 = FALSE) AND  ( TRUE ) AND  (x10 = FALSE) AND  (t0.Q = TRUE) AND  ( TRUE )) THEN 
        cstate64 := 33; y2 := FALSE; y3 := FALSE; t0_start := FALSE;t1_start := FALSE; 
    ELSIF ((x2 = FALSE) AND  ( TRUE ) AND  (x10 = TRUE) AND  (t0.Q = FALSE) AND  ( TRUE )) THEN 
        cstate64 := 20; y2 := FALSE; y3 := FALSE; t0_start := FALSE;t1_start := FALSE; 
    ELSIF ((x2 = FALSE) AND  ( TRUE ) AND  (x10 = TRUE) AND  (t0.Q = TRUE) AND  ( TRUE )) THEN 
        cstate64 := 33; y2 := FALSE; y3 := FALSE; t0_start := FALSE;t1_start := FALSE; 
    ELSIF ((x2 = TRUE) AND  ( TRUE ) AND  (x10 = FALSE) AND  (t0.Q = FALSE) AND  (t1.Q = FALSE)) THEN 
        cstate64 := 84; y2 := TRUE; y3 := FALSE; t0_start := FALSE;t1_start := FALSE; 
    ELSIF ((x2 = TRUE) AND  ( TRUE ) AND  (x10 = FALSE) AND  (t0.Q = FALSE) AND  (t1.Q = TRUE)) THEN 
        cstate64 := 84; y2 := TRUE; y3 := FALSE; t0_start := FALSE;t1_start := FALSE; 
    ELSIF ((x2 = TRUE) AND  ( TRUE ) AND  ( TRUE ) AND  (t0.Q = TRUE) AND  ( TRUE )) THEN 
        cstate64 := 65; y2 := FALSE; y3 := FALSE; t0_start := FALSE;t1_start := FALSE; 
    ELSIF ((x2 = TRUE) AND  ( TRUE ) AND  (x10 = TRUE) AND  (t0.Q = FALSE) AND  ( TRUE )) THEN 
        cstate64 := 52; y2 := FALSE; y3 := FALSE; t0_start := FALSE;t1_start := FALSE; 
    END_IF;
86:
    IF ((x2 = FALSE) AND  ( TRUE ) AND  (x10 = FALSE) AND  (t0.Q = FALSE) AND  (t1.Q = FALSE)) THEN 
        cstate64 := 106; y2 := TRUE; y3 := TRUE; t0_start := FALSE;t1_start := FALSE; 
    ELSIF ((x2 = FALSE) AND  ( TRUE ) AND  (x10 = FALSE) AND  (t0.Q = FALSE) AND  (t1.Q = TRUE)) THEN 
        cstate64 := 100; y2 := TRUE; y3 := FALSE; t0_start := FALSE;t1_start := FALSE; 
    ELSIF ((x2 = FALSE) AND  ( TRUE ) AND  (x10 = FALSE) AND  (t0.Q = TRUE) AND  (t1.Q = FALSE)) THEN 
        cstate64 := 37; y2 := FALSE; y3 := TRUE; t0_start := FALSE;t1_start := FALSE; 
    ELSIF ((x2 = FALSE) AND  ( TRUE ) AND  (x10 = FALSE) AND  (t0.Q = TRUE) AND  (t1.Q = TRUE)) THEN 
        cstate64 := 33; y2 := FALSE; y3 := FALSE; t0_start := FALSE;t1_start := FALSE; 
    ELSIF ((x2 = FALSE) AND  ( TRUE ) AND  (x10 = TRUE) AND  (t0.Q = FALSE) AND  (t1.Q = FALSE)) THEN 
        cstate64 := 19; y2 := FALSE; y3 := FALSE; t0_start := FALSE;t1_start := FALSE; 
    ELSIF ((x2 = FALSE) AND  ( TRUE ) AND  (x10 = TRUE) AND  (t0.Q = FALSE) AND  (t1.Q = TRUE)) THEN 
        cstate64 := 20; y2 := FALSE; y3 := FALSE; t0_start := FALSE;t1_start := FALSE; 
    ELSIF ((x2 = FALSE) AND  ( TRUE ) AND  (x10 = TRUE) AND  (t0.Q = TRUE) AND  (t1.Q = FALSE)) THEN 
        cstate64 := 34; y2 := FALSE; y3 := FALSE; t0_start := FALSE;t1_start := FALSE; 
    ELSIF ((x2 = FALSE) AND  ( TRUE ) AND  (x10 = TRUE) AND  (t0.Q = TRUE) AND  (t1.Q = TRUE)) THEN 
        cstate64 := 33; y2 := FALSE; y3 := FALSE; t0_start := FALSE;t1_start := FALSE; 
    ELSIF ((x2 = TRUE) AND  ( TRUE ) AND  (x10 = FALSE) AND  (t0.Q = FALSE) AND  (t1.Q = FALSE)) THEN 
        cstate64 := 90; y2 := TRUE; y3 := TRUE; t0_start := FALSE;t1_start := FALSE; 
    ELSIF ((x2 = TRUE) AND  ( TRUE ) AND  (x10 = FALSE) AND  (t0.Q = FALSE) AND  (t1.Q = TRUE)) THEN 
        cstate64 := 84; y2 := TRUE; y3 := FALSE; t0_start := FALSE;t1_start := FALSE; 
    ELSIF ((x2 = TRUE) AND  ( TRUE ) AND  (x10 = FALSE) AND  (t0.Q = TRUE) AND  (t1.Q = FALSE)) THEN 
        cstate64 := 69; y2 := FALSE; y3 := TRUE; t0_start := FALSE;t1_start := FALSE; 
    ELSIF ((x2 = TRUE) AND  ( TRUE ) AND  ( TRUE ) AND  (t0.Q = TRUE) AND  (t1.Q = TRUE)) THEN 
        cstate64 := 65; y2 := FALSE; y3 := FALSE; t0_start := FALSE;t1_start := FALSE; 
    ELSIF ((x2 = TRUE) AND  ( TRUE ) AND  (x10 = TRUE) AND  (t0.Q = FALSE) AND  (t1.Q = FALSE)) THEN 
        cstate64 := 51; y2 := FALSE; y3 := FALSE; t0_start := FALSE;t1_start := FALSE; 
    ELSIF ((x2 = TRUE) AND  ( TRUE ) AND  (x10 = TRUE) AND  (t0.Q = FALSE) AND  (t1.Q = TRUE)) THEN 
        cstate64 := 52; y2 := FALSE; y3 := FALSE; t0_start := FALSE;t1_start := FALSE; 
    ELSIF ((x2 = TRUE) AND  ( TRUE ) AND  (x10 = TRUE) AND  (t0.Q = TRUE) AND  (t1.Q = FALSE)) THEN 
        cstate64 := 66; y2 := FALSE; y3 := FALSE; t0_start := FALSE;t1_start := FALSE; 
    END_IF;
99:
    IF ((x2 = FALSE) AND  ( TRUE ) AND  (x10 = FALSE) AND  (t0.Q = FALSE) AND  (t1.Q = FALSE)) THEN 
        cstate64 := 99; y2 := TRUE; y3 := FALSE; t0_start := FALSE;t1_start := FALSE; 
    ELSIF ((x2 = FALSE) AND  ( TRUE ) AND  (x10 = FALSE) AND  (t0.Q = FALSE) AND  (t1.Q = TRUE)) THEN 
        cstate64 := 100; y2 := TRUE; y3 := FALSE; t0_start := FALSE;t1_start := FALSE; 
    ELSIF ((x2 = FALSE) AND  ( TRUE ) AND  (x10 = FALSE) AND  (t0.Q = TRUE) AND  ( TRUE )) THEN 
        cstate64 := 37; y2 := FALSE; y3 := TRUE; t0_start := FALSE;t1_start := TRUE; t1_up := FALSE; 
    ELSIF ((x2 = FALSE) AND  ( TRUE ) AND  (x10 = TRUE) AND  (t0.Q = FALSE) AND  (t1.Q = FALSE)) THEN 
        cstate64 := 19; y2 := FALSE; y3 := FALSE; t0_start := FALSE;t1_start := FALSE; 
    ELSIF ((x2 = FALSE) AND  ( TRUE ) AND  (x10 = TRUE) AND  (t0.Q = FALSE) AND  (t1.Q = TRUE)) THEN 
        cstate64 := 20; y2 := FALSE; y3 := FALSE; t0_start := FALSE;t1_start := FALSE; 
    ELSIF ((x2 = FALSE) AND  ( TRUE ) AND  (x10 = TRUE) AND  (t0.Q = TRUE) AND  (t1.Q = FALSE)) THEN 
        cstate64 := 34; y2 := FALSE; y3 := FALSE; t0_start := FALSE;t1_start := FALSE; 
    ELSIF ((x2 = FALSE) AND  ( TRUE ) AND  (x10 = TRUE) AND  (t0.Q = TRUE) AND  (t1.Q = TRUE)) THEN 
        cstate64 := 33; y2 := FALSE; y3 := FALSE; t0_start := FALSE;t1_start := FALSE; 
    ELSIF ((x2 = TRUE) AND  ( TRUE ) AND  (x10 = FALSE) AND  (t0.Q = FALSE) AND  (t1.Q = FALSE)) THEN 
        cstate64 := 83; y2 := TRUE; y3 := FALSE; t0_start := TRUE; t0_up := FALSE;t1_start := FALSE; 
    ELSIF ((x2 = TRUE) AND  ( TRUE ) AND  (x10 = FALSE) AND  (t0.Q = FALSE) AND  (t1.Q = TRUE)) THEN 
        cstate64 := 84; y2 := TRUE; y3 := FALSE; t0_start := TRUE; t0_up := FALSE;t1_start := FALSE; 
    ELSIF ((x2 = TRUE) AND  ( TRUE ) AND  (x10 = FALSE) AND  (t0.Q = TRUE) AND  ( TRUE )) THEN 
        cstate64 := 86; y2 := TRUE; y3 := TRUE; t0_start := TRUE; t0_up := FALSE;t1_start := TRUE; t1_up := FALSE; 
    ELSIF ((x2 = TRUE) AND  ( TRUE ) AND  (x10 = TRUE) AND  (t0.Q = FALSE) AND  (t1.Q = FALSE)) THEN 
        cstate64 := 51; y2 := FALSE; y3 := FALSE; t0_start := FALSE;t1_start := FALSE; 
    ELSIF ((x2 = TRUE) AND  ( TRUE ) AND  (x10 = TRUE) AND  (t0.Q = FALSE) AND  (t1.Q = TRUE)) THEN 
        cstate64 := 52; y2 := FALSE; y3 := FALSE; t0_start := FALSE;t1_start := FALSE; 
    ELSIF ((x2 = TRUE) AND  ( TRUE ) AND  (x10 = TRUE) AND  (t0.Q = TRUE) AND  (t1.Q = FALSE)) THEN 
        cstate64 := 66; y2 := FALSE; y3 := FALSE; t0_start := FALSE;t1_start := FALSE; 
    ELSIF ((x2 = TRUE) AND  ( TRUE ) AND  (x10 = TRUE) AND  (t0.Q = TRUE) AND  (t1.Q = TRUE)) THEN 
        cstate64 := 65; y2 := FALSE; y3 := FALSE; t0_start := FALSE;t1_start := FALSE; 
    END_IF;
87:
    IF ((x2 = FALSE) AND  ( TRUE ) AND  (x10 = FALSE) AND  (t0.Q = FALSE) AND  (t1.Q = FALSE)) THEN 
        cstate64 := 107; y2 := TRUE; y3 := TRUE; t0_start := FALSE;t1_start := FALSE; 
    ELSIF ((x2 = FALSE) AND  ( TRUE ) AND  (x10 = FALSE) AND  (t0.Q = FALSE) AND  (t1.Q = TRUE)) THEN 
        cstate64 := 100; y2 := TRUE; y3 := FALSE; t0_start := FALSE;t1_start := FALSE; 
    ELSIF ((x2 = FALSE) AND  ( TRUE ) AND  (x10 = FALSE) AND  (t0.Q = TRUE) AND  (t1.Q = FALSE)) THEN 
        cstate64 := 40; y2 := FALSE; y3 := TRUE; t0_start := FALSE;t1_start := FALSE; 
    ELSIF ((x2 = FALSE) AND  ( TRUE ) AND  (x10 = FALSE) AND  (t0.Q = TRUE) AND  (t1.Q = TRUE)) THEN 
        cstate64 := 33; y2 := FALSE; y3 := FALSE; t0_start := FALSE;t1_start := FALSE; 
    ELSIF ((x2 = FALSE) AND  ( TRUE ) AND  (x10 = TRUE) AND  (t0.Q = FALSE) AND  (t1.Q = FALSE)) THEN 
        cstate64 := 19; y2 := FALSE; y3 := FALSE; t0_start := FALSE;t1_start := FALSE; 
    ELSIF ((x2 = FALSE) AND  ( TRUE ) AND  (x10 = TRUE) AND  (t0.Q = FALSE) AND  (t1.Q = TRUE)) THEN 
        cstate64 := 20; y2 := FALSE; y3 := FALSE; t0_start := FALSE;t1_start := FALSE; 
    ELSIF ((x2 = FALSE) AND  ( TRUE ) AND  (x10 = TRUE) AND  (t0.Q = TRUE) AND  (t1.Q = FALSE)) THEN 
        cstate64 := 34; y2 := FALSE; y3 := FALSE; t0_start := FALSE;t1_start := FALSE; 
    ELSIF ((x2 = FALSE) AND  ( TRUE ) AND  (x10 = TRUE) AND  (t0.Q = TRUE) AND  (t1.Q = TRUE)) THEN 
        cstate64 := 33; y2 := FALSE; y3 := FALSE; t0_start := FALSE;t1_start := FALSE; 
    ELSIF ((x2 = TRUE) AND  ( TRUE ) AND  (x10 = FALSE) AND  (t0.Q = FALSE) AND  (t1.Q = FALSE)) THEN 
        cstate64 := 91; y2 := TRUE; y3 := TRUE; t0_start := FALSE;t1_start := FALSE; 
    ELSIF ((x2 = TRUE) AND  ( TRUE ) AND  (x10 = FALSE) AND  (t0.Q = FALSE) AND  (t1.Q = TRUE)) THEN 
        cstate64 := 84; y2 := TRUE; y3 := FALSE; t0_start := FALSE;t1_start := FALSE; 
    ELSIF ((x2 = TRUE) AND  ( TRUE ) AND  (x10 = FALSE) AND  (t0.Q = TRUE) AND  (t1.Q = FALSE)) THEN 
        cstate64 := 72; y2 := FALSE; y3 := TRUE; t0_start := FALSE;t1_start := FALSE; 
    ELSIF ((x2 = TRUE) AND  ( TRUE ) AND  ( TRUE ) AND  (t0.Q = TRUE) AND  (t1.Q = TRUE)) THEN 
        cstate64 := 65; y2 := FALSE; y3 := FALSE; t0_start := FALSE;t1_start := FALSE; 
    ELSIF ((x2 = TRUE) AND  ( TRUE ) AND  (x10 = TRUE) AND  (t0.Q = FALSE) AND  (t1.Q = FALSE)) THEN 
        cstate64 := 51; y2 := FALSE; y3 := FALSE; t0_start := FALSE;t1_start := FALSE; 
    ELSIF ((x2 = TRUE) AND  ( TRUE ) AND  (x10 = TRUE) AND  (t0.Q = FALSE) AND  (t1.Q = TRUE)) THEN 
        cstate64 := 52; y2 := FALSE; y3 := FALSE; t0_start := FALSE;t1_start := FALSE; 
    ELSIF ((x2 = TRUE) AND  ( TRUE ) AND  (x10 = TRUE) AND  (t0.Q = TRUE) AND  (t1.Q = FALSE)) THEN 
        cstate64 := 66; y2 := FALSE; y3 := FALSE; t0_start := FALSE;t1_start := FALSE; 
    END_IF;
100:
    IF ((x2 = FALSE) AND  ( TRUE ) AND  (x10 = FALSE) AND  (t0.Q = FALSE) AND  (t1.Q = FALSE)) THEN 
        cstate64 := 100; y2 := TRUE; y3 := FALSE; t0_start := FALSE;t1_start := FALSE; 
    ELSIF ((x2 = FALSE) AND  ( TRUE ) AND  (x10 = FALSE) AND  (t0.Q = FALSE) AND  (t1.Q = TRUE)) THEN 
        cstate64 := 100; y2 := TRUE; y3 := FALSE; t0_start := FALSE;t1_start := FALSE; 
    ELSIF ((x2 = FALSE) AND  ( TRUE ) AND  (x10 = FALSE) AND  (t0.Q = TRUE) AND  ( TRUE )) THEN 
        cstate64 := 40; y2 := FALSE; y3 := TRUE; t0_start := FALSE;t1_start := TRUE; t1_up := FALSE; 
    ELSIF ((x2 = FALSE) AND  ( TRUE ) AND  (x10 = TRUE) AND  (t0.Q = FALSE) AND  ( TRUE )) THEN 
        cstate64 := 20; y2 := FALSE; y3 := FALSE; t0_start := FALSE;t1_start := FALSE; 
    ELSIF ((x2 = FALSE) AND  ( TRUE ) AND  (x10 = TRUE) AND  (t0.Q = TRUE) AND  ( TRUE )) THEN 
        cstate64 := 33; y2 := FALSE; y3 := FALSE; t0_start := FALSE;t1_start := FALSE; 
    ELSIF ((x2 = TRUE) AND  ( TRUE ) AND  (x10 = FALSE) AND  (t0.Q = FALSE) AND  (t1.Q = FALSE)) THEN 
        cstate64 := 84; y2 := TRUE; y3 := FALSE; t0_start := TRUE; t0_up := FALSE;t1_start := FALSE; 
    ELSIF ((x2 = TRUE) AND  ( TRUE ) AND  (x10 = FALSE) AND  (t0.Q = FALSE) AND  (t1.Q = TRUE)) THEN 
        cstate64 := 84; y2 := TRUE; y3 := FALSE; t0_start := TRUE; t0_up := FALSE;t1_start := FALSE; 
    ELSIF ((x2 = TRUE) AND  ( TRUE ) AND  (x10 = FALSE) AND  (t0.Q = TRUE) AND  ( TRUE )) THEN 
        cstate64 := 87; y2 := TRUE; y3 := TRUE; t0_start := TRUE; t0_up := FALSE;t1_start := TRUE; t1_up := FALSE; 
    ELSIF ((x2 = TRUE) AND  ( TRUE ) AND  (x10 = TRUE) AND  (t0.Q = FALSE) AND  ( TRUE )) THEN 
        cstate64 := 52; y2 := FALSE; y3 := FALSE; t0_start := FALSE;t1_start := FALSE; 
    ELSIF ((x2 = TRUE) AND  ( TRUE ) AND  (x10 = TRUE) AND  (t0.Q = TRUE) AND  ( TRUE )) THEN 
        cstate64 := 65; y2 := FALSE; y3 := FALSE; t0_start := FALSE;t1_start := FALSE; 
    END_IF;
84:
    IF ((x2 = FALSE) AND  ( TRUE ) AND  (x10 = FALSE) AND  (t0.Q = FALSE) AND  (t1.Q = FALSE)) THEN 
        cstate64 := 100; y2 := TRUE; y3 := FALSE; t0_start := FALSE;t1_start := FALSE; 
    ELSIF ((x2 = FALSE) AND  ( TRUE ) AND  (x10 = FALSE) AND  (t0.Q = FALSE) AND  (t1.Q = TRUE)) THEN 
        cstate64 := 100; y2 := TRUE; y3 := FALSE; t0_start := FALSE;t1_start := FALSE; 
    ELSIF ((x2 = FALSE) AND  ( TRUE ) AND  (x10 = FALSE) AND  (t0.Q = TRUE) AND  ( TRUE )) THEN 
        cstate64 := 40; y2 := FALSE; y3 := TRUE; t0_start := FALSE;t1_start := TRUE; t1_up := FALSE; 
    ELSIF ((x2 = FALSE) AND  ( TRUE ) AND  (x10 = TRUE) AND  (t0.Q = FALSE) AND  ( TRUE )) THEN 
        cstate64 := 20; y2 := FALSE; y3 := FALSE; t0_start := FALSE;t1_start := FALSE; 
    ELSIF ((x2 = FALSE) AND  ( TRUE ) AND  (x10 = TRUE) AND  (t0.Q = TRUE) AND  ( TRUE )) THEN 
        cstate64 := 33; y2 := FALSE; y3 := FALSE; t0_start := FALSE;t1_start := FALSE; 
    ELSIF ((x2 = TRUE) AND  ( TRUE ) AND  (x10 = FALSE) AND  (t0.Q = FALSE) AND  (t1.Q = FALSE)) THEN 
        cstate64 := 84; y2 := TRUE; y3 := FALSE; t0_start := FALSE;t1_start := FALSE; 
    ELSIF ((x2 = TRUE) AND  ( TRUE ) AND  (x10 = FALSE) AND  (t0.Q = FALSE) AND  (t1.Q = TRUE)) THEN 
        cstate64 := 84; y2 := TRUE; y3 := FALSE; t0_start := FALSE;t1_start := FALSE; 
    ELSIF ((x2 = TRUE) AND  ( TRUE ) AND  (x10 = FALSE) AND  (t0.Q = TRUE) AND  ( TRUE )) THEN 
        cstate64 := 72; y2 := FALSE; y3 := TRUE; t0_start := FALSE;t1_start := TRUE; t1_up := FALSE; 
    ELSIF ((x2 = TRUE) AND  ( TRUE ) AND  (x10 = TRUE) AND  (t0.Q = FALSE) AND  ( TRUE )) THEN 
        cstate64 := 52; y2 := FALSE; y3 := FALSE; t0_start := FALSE;t1_start := FALSE; 
    ELSIF ((x2 = TRUE) AND  ( TRUE ) AND  (x10 = TRUE) AND  (t0.Q = TRUE) AND  ( TRUE )) THEN 
        cstate64 := 65; y2 := FALSE; y3 := FALSE; t0_start := FALSE;t1_start := FALSE; 
    END_IF;
67:
    IF ((x2 = FALSE) AND  ( TRUE ) AND  ( TRUE ) AND  (t0.Q = FALSE) AND  (t1.Q = FALSE)) THEN 
        cstate64 := 35; y2 := FALSE; y3 := FALSE; t0_start := FALSE;t1_start := FALSE; 
    ELSIF ((x2 = FALSE) AND  ( TRUE ) AND  (x10 = FALSE) AND  (t0.Q = FALSE) AND  (t1.Q = TRUE)) THEN 
        cstate64 := 36; y2 := FALSE; y3 := FALSE; t0_start := FALSE;t1_start := FALSE; 
    ELSIF ((x2 = FALSE) AND  ( TRUE ) AND  (x10 = FALSE) AND  (t0.Q = TRUE) AND  ( TRUE )) THEN 
        cstate64 := 37; y2 := FALSE; y3 := TRUE; t0_start := FALSE;t1_start := TRUE; t1_up := FALSE; 
    ELSIF ((x2 = FALSE) AND  ( TRUE ) AND  (x10 = TRUE) AND  (t0.Q = FALSE) AND  (t1.Q = TRUE)) THEN 
        cstate64 := 36; y2 := FALSE; y3 := FALSE; t0_start := FALSE;t1_start := FALSE; 
    ELSIF ((x2 = FALSE) AND  ( TRUE ) AND  (x10 = TRUE) AND  (t0.Q = TRUE) AND  (t1.Q = FALSE)) THEN 
        cstate64 := 34; y2 := FALSE; y3 := FALSE; t0_start := FALSE;t1_start := FALSE; 
    ELSIF ((x2 = FALSE) AND  ( TRUE ) AND  (x10 = TRUE) AND  (t0.Q = TRUE) AND  (t1.Q = TRUE)) THEN 
        cstate64 := 33; y2 := FALSE; y3 := FALSE; t0_start := FALSE;t1_start := FALSE; 
    ELSIF ((x2 = TRUE) AND  ( TRUE ) AND  ( TRUE ) AND  (t0.Q = FALSE) AND  (t1.Q = FALSE)) THEN 
        cstate64 := 67; y2 := FALSE; y3 := FALSE; t0_start := FALSE;t1_start := FALSE; 
    ELSIF ((x2 = TRUE) AND  ( TRUE ) AND  (x10 = FALSE) AND  (t0.Q = FALSE) AND  (t1.Q = TRUE)) THEN 
        cstate64 := 68; y2 := FALSE; y3 := FALSE; t0_start := FALSE;t1_start := FALSE; 
    ELSIF ((x2 = TRUE) AND  ( TRUE ) AND  (x10 = FALSE) AND  (t0.Q = TRUE) AND  ( TRUE )) THEN 
        cstate64 := 69; y2 := FALSE; y3 := TRUE; t0_start := FALSE;t1_start := TRUE; t1_up := FALSE; 
    ELSIF ((x2 = TRUE) AND  ( TRUE ) AND  (x10 = TRUE) AND  (t0.Q = FALSE) AND  (t1.Q = TRUE)) THEN 
        cstate64 := 68; y2 := FALSE; y3 := FALSE; t0_start := FALSE;t1_start := FALSE; 
    ELSIF ((x2 = TRUE) AND  ( TRUE ) AND  (x10 = TRUE) AND  (t0.Q = TRUE) AND  (t1.Q = FALSE)) THEN 
        cstate64 := 66; y2 := FALSE; y3 := FALSE; t0_start := FALSE;t1_start := FALSE; 
    ELSIF ((x2 = TRUE) AND  ( TRUE ) AND  (x10 = TRUE) AND  (t0.Q = TRUE) AND  (t1.Q = TRUE)) THEN 
        cstate64 := 65; y2 := FALSE; y3 := FALSE; t0_start := FALSE;t1_start := FALSE; 
    END_IF;
66:
    IF ((x2 = FALSE) AND  ( TRUE ) AND  ( TRUE ) AND  (t0.Q = FALSE) AND  (t1.Q = FALSE)) THEN 
        cstate64 := 35; y2 := FALSE; y3 := FALSE; t0_start := FALSE;t1_start := FALSE; 
    ELSIF ((x2 = FALSE) AND  ( TRUE ) AND  (x10 = FALSE) AND  (t0.Q = FALSE) AND  (t1.Q = TRUE)) THEN 
        cstate64 := 36; y2 := FALSE; y3 := FALSE; t0_start := FALSE;t1_start := FALSE; 
    ELSIF ((x2 = FALSE) AND  ( TRUE ) AND  (x10 = FALSE) AND  (t0.Q = TRUE) AND  (t1.Q = FALSE)) THEN 
        cstate64 := 34; y2 := FALSE; y3 := FALSE; t0_start := FALSE;t1_start := FALSE; 
    ELSIF ((x2 = FALSE) AND  ( TRUE ) AND  (x10 = FALSE) AND  (t0.Q = TRUE) AND  (t1.Q = TRUE)) THEN 
        cstate64 := 33; y2 := FALSE; y3 := FALSE; t0_start := FALSE;t1_start := FALSE; 
    ELSIF ((x2 = FALSE) AND  ( TRUE ) AND  (x10 = TRUE) AND  (t0.Q = FALSE) AND  (t1.Q = TRUE)) THEN 
        cstate64 := 36; y2 := FALSE; y3 := FALSE; t0_start := FALSE;t1_start := FALSE; 
    ELSIF ((x2 = FALSE) AND  ( TRUE ) AND  (x10 = TRUE) AND  (t0.Q = TRUE) AND  (t1.Q = FALSE)) THEN 
        cstate64 := 34; y2 := FALSE; y3 := FALSE; t0_start := FALSE;t1_start := FALSE; 
    ELSIF ((x2 = FALSE) AND  ( TRUE ) AND  (x10 = TRUE) AND  (t0.Q = TRUE) AND  (t1.Q = TRUE)) THEN 
        cstate64 := 33; y2 := FALSE; y3 := FALSE; t0_start := FALSE;t1_start := FALSE; 
    ELSIF ((x2 = TRUE) AND  ( TRUE ) AND  ( TRUE ) AND  (t0.Q = FALSE) AND  (t1.Q = FALSE)) THEN 
        cstate64 := 67; y2 := FALSE; y3 := FALSE; t0_start := FALSE;t1_start := FALSE; 
    ELSIF ((x2 = TRUE) AND  ( TRUE ) AND  (x10 = FALSE) AND  (t0.Q = FALSE) AND  (t1.Q = TRUE)) THEN 
        cstate64 := 68; y2 := FALSE; y3 := FALSE; t0_start := FALSE;t1_start := FALSE; 
    ELSIF ((x2 = TRUE) AND  ( TRUE ) AND  ( TRUE ) AND  (t0.Q = TRUE) AND  (t1.Q = FALSE)) THEN 
        cstate64 := 66; y2 := FALSE; y3 := FALSE; t0_start := FALSE;t1_start := FALSE; 
    ELSIF ((x2 = TRUE) AND  ( TRUE ) AND  ( TRUE ) AND  (t0.Q = TRUE) AND  (t1.Q = TRUE)) THEN 
        cstate64 := 65; y2 := FALSE; y3 := FALSE; t0_start := FALSE;t1_start := FALSE; 
    ELSIF ((x2 = TRUE) AND  ( TRUE ) AND  (x10 = TRUE) AND  (t0.Q = FALSE) AND  (t1.Q = TRUE)) THEN 
        cstate64 := 68; y2 := FALSE; y3 := FALSE; t0_start := FALSE;t1_start := FALSE; 
    END_IF;
69:
    IF ((x2 = FALSE) AND  ( TRUE ) AND  (x10 = FALSE) AND  (t0.Q = FALSE) AND  (t1.Q = FALSE)) THEN 
        cstate64 := 41; y2 := FALSE; y3 := TRUE; t0_start := FALSE;t1_start := FALSE; 
    ELSIF ((x2 = FALSE) AND  ( TRUE ) AND  (x10 = FALSE) AND  (t0.Q = FALSE) AND  (t1.Q = TRUE)) THEN 
        cstate64 := 36; y2 := FALSE; y3 := FALSE; t0_start := FALSE;t1_start := FALSE; 
    ELSIF ((x2 = FALSE) AND  ( TRUE ) AND  (x10 = FALSE) AND  (t0.Q = TRUE) AND  (t1.Q = FALSE)) THEN 
        cstate64 := 37; y2 := FALSE; y3 := TRUE; t0_start := FALSE;t1_start := FALSE; 
    ELSIF ((x2 = FALSE) AND  ( TRUE ) AND  (x10 = FALSE) AND  (t0.Q = TRUE) AND  (t1.Q = TRUE)) THEN 
        cstate64 := 33; y2 := FALSE; y3 := FALSE; t0_start := FALSE;t1_start := FALSE; 
    ELSIF ((x2 = FALSE) AND  ( TRUE ) AND  (x10 = TRUE) AND  (t0.Q = FALSE) AND  (t1.Q = FALSE)) THEN 
        cstate64 := 35; y2 := FALSE; y3 := FALSE; t0_start := FALSE;t1_start := FALSE; 
    ELSIF ((x2 = FALSE) AND  ( TRUE ) AND  (x10 = TRUE) AND  (t0.Q = FALSE) AND  (t1.Q = TRUE)) THEN 
        cstate64 := 36; y2 := FALSE; y3 := FALSE; t0_start := FALSE;t1_start := FALSE; 
    ELSIF ((x2 = FALSE) AND  ( TRUE ) AND  (x10 = TRUE) AND  (t0.Q = TRUE) AND  (t1.Q = FALSE)) THEN 
        cstate64 := 34; y2 := FALSE; y3 := FALSE; t0_start := FALSE;t1_start := FALSE; 
    ELSIF ((x2 = FALSE) AND  ( TRUE ) AND  (x10 = TRUE) AND  (t0.Q = TRUE) AND  (t1.Q = TRUE)) THEN 
        cstate64 := 33; y2 := FALSE; y3 := FALSE; t0_start := FALSE;t1_start := FALSE; 
    ELSIF ((x2 = TRUE) AND  ( TRUE ) AND  (x10 = FALSE) AND  (t0.Q = FALSE) AND  (t1.Q = FALSE)) THEN 
        cstate64 := 73; y2 := FALSE; y3 := TRUE; t0_start := FALSE;t1_start := FALSE; 
    ELSIF ((x2 = TRUE) AND  ( TRUE ) AND  (x10 = FALSE) AND  (t0.Q = FALSE) AND  (t1.Q = TRUE)) THEN 
        cstate64 := 68; y2 := FALSE; y3 := FALSE; t0_start := FALSE;t1_start := FALSE; 
    ELSIF ((x2 = TRUE) AND  ( TRUE ) AND  (x10 = FALSE) AND  (t0.Q = TRUE) AND  (t1.Q = FALSE)) THEN 
        cstate64 := 69; y2 := FALSE; y3 := TRUE; t0_start := FALSE;t1_start := FALSE; 
    ELSIF ((x2 = TRUE) AND  ( TRUE ) AND  ( TRUE ) AND  (t0.Q = TRUE) AND  (t1.Q = TRUE)) THEN 
        cstate64 := 65; y2 := FALSE; y3 := FALSE; t0_start := FALSE;t1_start := FALSE; 
    ELSIF ((x2 = TRUE) AND  ( TRUE ) AND  (x10 = TRUE) AND  (t0.Q = FALSE) AND  (t1.Q = FALSE)) THEN 
        cstate64 := 67; y2 := FALSE; y3 := FALSE; t0_start := FALSE;t1_start := FALSE; 
    ELSIF ((x2 = TRUE) AND  ( TRUE ) AND  (x10 = TRUE) AND  (t0.Q = FALSE) AND  (t1.Q = TRUE)) THEN 
        cstate64 := 68; y2 := FALSE; y3 := FALSE; t0_start := FALSE;t1_start := FALSE; 
    ELSIF ((x2 = TRUE) AND  ( TRUE ) AND  (x10 = TRUE) AND  (t0.Q = TRUE) AND  (t1.Q = FALSE)) THEN 
        cstate64 := 66; y2 := FALSE; y3 := FALSE; t0_start := FALSE;t1_start := FALSE; 
    END_IF;
68:
    IF ((x2 = FALSE) AND  ( TRUE ) AND  (x10 = FALSE) AND  (t0.Q = FALSE) AND  (t1.Q = FALSE)) OR ((x2 = FALSE) AND  ( TRUE ) AND  (x10 = TRUE) AND  (t0.Q = FALSE) AND  ( TRUE )) THEN 
        cstate64 := 36; y2 := FALSE; y3 := FALSE; t0_start := FALSE;t1_start := FALSE; 
    ELSIF ((x2 = FALSE) AND  ( TRUE ) AND  (x10 = FALSE) AND  (t0.Q = FALSE) AND  (t1.Q = TRUE)) THEN 
        cstate64 := 36; y2 := FALSE; y3 := FALSE; t0_start := FALSE;t1_start := FALSE; 
    ELSIF ((x2 = FALSE) AND  ( TRUE ) AND  (x10 = FALSE) AND  (t0.Q = TRUE) AND  ( TRUE )) THEN 
        cstate64 := 40; y2 := FALSE; y3 := TRUE; t0_start := FALSE;t1_start := TRUE; t1_up := FALSE; 
    ELSIF ((x2 = FALSE) AND  ( TRUE ) AND  (x10 = TRUE) AND  (t0.Q = TRUE) AND  ( TRUE )) THEN 
        cstate64 := 33; y2 := FALSE; y3 := FALSE; t0_start := FALSE;t1_start := FALSE; 
    ELSIF ((x2 = TRUE) AND  ( TRUE ) AND  (x10 = FALSE) AND  (t0.Q = FALSE) AND  (t1.Q = FALSE)) OR ((x2 = TRUE) AND  ( TRUE ) AND  (x10 = TRUE) AND  (t0.Q = FALSE) AND  ( TRUE )) THEN 
        cstate64 := 68; y2 := FALSE; y3 := FALSE; t0_start := FALSE;t1_start := FALSE; 
    ELSIF ((x2 = TRUE) AND  ( TRUE ) AND  (x10 = FALSE) AND  (t0.Q = FALSE) AND  (t1.Q = TRUE)) THEN 
        cstate64 := 68; y2 := FALSE; y3 := FALSE; t0_start := FALSE;t1_start := FALSE; 
    ELSIF ((x2 = TRUE) AND  ( TRUE ) AND  (x10 = FALSE) AND  (t0.Q = TRUE) AND  ( TRUE )) THEN 
        cstate64 := 72; y2 := FALSE; y3 := TRUE; t0_start := FALSE;t1_start := TRUE; t1_up := FALSE; 
    ELSIF ((x2 = TRUE) AND  ( TRUE ) AND  (x10 = TRUE) AND  (t0.Q = TRUE) AND  ( TRUE )) THEN 
        cstate64 := 65; y2 := FALSE; y3 := FALSE; t0_start := FALSE;t1_start := FALSE; 
    END_IF;
44:
    IF ((x2 = FALSE) AND  ( TRUE ) AND  (x10 = FALSE) AND  (t0.Q = FALSE) AND  (t1.Q = FALSE)) THEN 
        cstate64 := 44; y2 := FALSE; y3 := TRUE; t0_start := FALSE;t1_start := FALSE; 
    ELSIF ((x2 = FALSE) AND  ( TRUE ) AND  (x10 = FALSE) AND  (t0.Q = FALSE) AND  (t1.Q = TRUE)) THEN 
        cstate64 := 36; y2 := FALSE; y3 := FALSE; t0_start := FALSE;t1_start := FALSE; 
    ELSIF ((x2 = FALSE) AND  ( TRUE ) AND  (x10 = FALSE) AND  (t0.Q = TRUE) AND  (t1.Q = FALSE)) THEN 
        cstate64 := 40; y2 := FALSE; y3 := TRUE; t0_start := FALSE;t1_start := TRUE; t1_up := FALSE; 
    ELSIF ((x2 = FALSE) AND  ( TRUE ) AND  (x10 = FALSE) AND  (t0.Q = TRUE) AND  (t1.Q = TRUE)) THEN 
        cstate64 := 37; y2 := FALSE; y3 := TRUE; t0_start := FALSE;t1_start := TRUE; t1_up := FALSE; 
    ELSIF ((x2 = FALSE) AND  ( TRUE ) AND  (x10 = TRUE) AND  (t0.Q = FALSE) AND  (t1.Q = FALSE)) THEN 
        cstate64 := 35; y2 := FALSE; y3 := FALSE; t0_start := FALSE;t1_start := FALSE; 
    ELSIF ((x2 = FALSE) AND  ( TRUE ) AND  (x10 = TRUE) AND  (t0.Q = FALSE) AND  (t1.Q = TRUE)) THEN 
        cstate64 := 36; y2 := FALSE; y3 := FALSE; t0_start := FALSE;t1_start := FALSE; 
    ELSIF ((x2 = FALSE) AND  ( TRUE ) AND  (x10 = TRUE) AND  (t0.Q = TRUE) AND  (t1.Q = FALSE)) THEN 
        cstate64 := 34; y2 := FALSE; y3 := FALSE; t0_start := FALSE;t1_start := FALSE; 
    ELSIF ((x2 = FALSE) AND  ( TRUE ) AND  (x10 = TRUE) AND  (t0.Q = TRUE) AND  (t1.Q = TRUE)) THEN 
        cstate64 := 33; y2 := FALSE; y3 := FALSE; t0_start := FALSE;t1_start := FALSE; 
    ELSIF ((x2 = TRUE) AND  ( TRUE ) AND  (x10 = FALSE) AND  (t0.Q = FALSE) AND  (t1.Q = FALSE)) THEN 
        cstate64 := 91; y2 := TRUE; y3 := TRUE; t0_start := TRUE; t0_up := FALSE;t1_start := FALSE; 
    ELSIF ((x2 = TRUE) AND  ( TRUE ) AND  (x10 = FALSE) AND  (t0.Q = FALSE) AND  (t1.Q = TRUE)) THEN 
        cstate64 := 84; y2 := TRUE; y3 := FALSE; t0_start := TRUE; t0_up := FALSE;t1_start := FALSE; 
    ELSIF ((x2 = TRUE) AND  ( TRUE ) AND  (x10 = FALSE) AND  (t0.Q = TRUE) AND  (t1.Q = FALSE)) THEN 
        cstate64 := 87; y2 := TRUE; y3 := TRUE; t0_start := TRUE; t0_up := FALSE;t1_start := TRUE; t1_up := FALSE; 
    ELSIF ((x2 = TRUE) AND  ( TRUE ) AND  (x10 = FALSE) AND  (t0.Q = TRUE) AND  (t1.Q = TRUE)) THEN 
        cstate64 := 86; y2 := TRUE; y3 := TRUE; t0_start := TRUE; t0_up := FALSE;t1_start := TRUE; t1_up := FALSE; 
    ELSIF ((x2 = TRUE) AND  ( TRUE ) AND  (x10 = TRUE) AND  (t0.Q = FALSE) AND  (t1.Q = FALSE)) THEN 
        cstate64 := 67; y2 := FALSE; y3 := FALSE; t0_start := FALSE;t1_start := FALSE; 
    ELSIF ((x2 = TRUE) AND  ( TRUE ) AND  (x10 = TRUE) AND  (t0.Q = FALSE) AND  (t1.Q = TRUE)) THEN 
        cstate64 := 68; y2 := FALSE; y3 := FALSE; t0_start := FALSE;t1_start := FALSE; 
    ELSIF ((x2 = TRUE) AND  ( TRUE ) AND  (x10 = TRUE) AND  (t0.Q = TRUE) AND  (t1.Q = FALSE)) THEN 
        cstate64 := 66; y2 := FALSE; y3 := FALSE; t0_start := FALSE;t1_start := FALSE; 
    ELSIF ((x2 = TRUE) AND  ( TRUE ) AND  (x10 = TRUE) AND  (t0.Q = TRUE) AND  (t1.Q = TRUE)) THEN 
        cstate64 := 65; y2 := FALSE; y3 := FALSE; t0_start := FALSE;t1_start := FALSE; 
    END_IF;
91:
    IF ((x2 = FALSE) AND  ( TRUE ) AND  (x10 = FALSE) AND  (t0.Q = FALSE) AND  (t1.Q = FALSE)) THEN 
        cstate64 := 107; y2 := TRUE; y3 := TRUE; t0_start := FALSE;t1_start := FALSE; 
    ELSIF ((x2 = FALSE) AND  ( TRUE ) AND  (x10 = FALSE) AND  (t0.Q = FALSE) AND  (t1.Q = TRUE)) THEN 
        cstate64 := 100; y2 := TRUE; y3 := FALSE; t0_start := FALSE;t1_start := FALSE; 
    ELSIF ((x2 = FALSE) AND  ( TRUE ) AND  (x10 = FALSE) AND  (t0.Q = TRUE) AND  (t1.Q = FALSE)) THEN 
        cstate64 := 40; y2 := FALSE; y3 := TRUE; t0_start := FALSE;t1_start := TRUE; t1_up := FALSE; 
    ELSIF ((x2 = FALSE) AND  ( TRUE ) AND  (x10 = FALSE) AND  (t0.Q = TRUE) AND  (t1.Q = TRUE)) THEN 
        cstate64 := 37; y2 := FALSE; y3 := TRUE; t0_start := FALSE;t1_start := TRUE; t1_up := FALSE; 
    ELSIF ((x2 = FALSE) AND  ( TRUE ) AND  (x10 = TRUE) AND  (t0.Q = FALSE) AND  (t1.Q = FALSE)) THEN 
        cstate64 := 19; y2 := FALSE; y3 := FALSE; t0_start := FALSE;t1_start := FALSE; 
    ELSIF ((x2 = FALSE) AND  ( TRUE ) AND  (x10 = TRUE) AND  (t0.Q = FALSE) AND  (t1.Q = TRUE)) THEN 
        cstate64 := 20; y2 := FALSE; y3 := FALSE; t0_start := FALSE;t1_start := FALSE; 
    ELSIF ((x2 = FALSE) AND  ( TRUE ) AND  (x10 = TRUE) AND  (t0.Q = TRUE) AND  (t1.Q = FALSE)) THEN 
        cstate64 := 34; y2 := FALSE; y3 := FALSE; t0_start := FALSE;t1_start := FALSE; 
    ELSIF ((x2 = FALSE) AND  ( TRUE ) AND  (x10 = TRUE) AND  (t0.Q = TRUE) AND  (t1.Q = TRUE)) THEN 
        cstate64 := 33; y2 := FALSE; y3 := FALSE; t0_start := FALSE;t1_start := FALSE; 
    ELSIF ((x2 = TRUE) AND  ( TRUE ) AND  (x10 = FALSE) AND  (t0.Q = FALSE) AND  (t1.Q = FALSE)) THEN 
        cstate64 := 91; y2 := TRUE; y3 := TRUE; t0_start := FALSE;t1_start := FALSE; 
    ELSIF ((x2 = TRUE) AND  ( TRUE ) AND  (x10 = FALSE) AND  (t0.Q = FALSE) AND  (t1.Q = TRUE)) THEN 
        cstate64 := 84; y2 := TRUE; y3 := FALSE; t0_start := FALSE;t1_start := FALSE; 
    ELSIF ((x2 = TRUE) AND  ( TRUE ) AND  (x10 = FALSE) AND  (t0.Q = TRUE) AND  (t1.Q = FALSE)) THEN 
        cstate64 := 72; y2 := FALSE; y3 := TRUE; t0_start := FALSE;t1_start := TRUE; t1_up := FALSE; 
    ELSIF ((x2 = TRUE) AND  ( TRUE ) AND  (x10 = FALSE) AND  (t0.Q = TRUE) AND  (t1.Q = TRUE)) THEN 
        cstate64 := 69; y2 := FALSE; y3 := TRUE; t0_start := FALSE;t1_start := TRUE; t1_up := FALSE; 
    ELSIF ((x2 = TRUE) AND  ( TRUE ) AND  (x10 = TRUE) AND  (t0.Q = FALSE) AND  (t1.Q = FALSE)) THEN 
        cstate64 := 51; y2 := FALSE; y3 := FALSE; t0_start := FALSE;t1_start := FALSE; 
    ELSIF ((x2 = TRUE) AND  ( TRUE ) AND  (x10 = TRUE) AND  (t0.Q = FALSE) AND  (t1.Q = TRUE)) THEN 
        cstate64 := 52; y2 := FALSE; y3 := FALSE; t0_start := FALSE;t1_start := FALSE; 
    ELSIF ((x2 = TRUE) AND  ( TRUE ) AND  (x10 = TRUE) AND  (t0.Q = TRUE) AND  (t1.Q = FALSE)) THEN 
        cstate64 := 66; y2 := FALSE; y3 := FALSE; t0_start := FALSE;t1_start := FALSE; 
    ELSIF ((x2 = TRUE) AND  ( TRUE ) AND  (x10 = TRUE) AND  (t0.Q = TRUE) AND  (t1.Q = TRUE)) THEN 
        cstate64 := 65; y2 := FALSE; y3 := FALSE; t0_start := FALSE;t1_start := FALSE; 
    END_IF;
90:
    IF ((x2 = FALSE) AND  ( TRUE ) AND  (x10 = FALSE) AND  (t0.Q = FALSE) AND  (t1.Q = FALSE)) THEN 
        cstate64 := 106; y2 := TRUE; y3 := TRUE; t0_start := FALSE;t1_start := FALSE; 
    ELSIF ((x2 = FALSE) AND  ( TRUE ) AND  (x10 = FALSE) AND  (t0.Q = FALSE) AND  (t1.Q = TRUE)) THEN 
        cstate64 := 100; y2 := TRUE; y3 := FALSE; t0_start := FALSE;t1_start := FALSE; 
    ELSIF ((x2 = FALSE) AND  ( TRUE ) AND  (x10 = FALSE) AND  (t0.Q = TRUE) AND  ( TRUE )) THEN 
        cstate64 := 37; y2 := FALSE; y3 := TRUE; t0_start := FALSE;t1_start := TRUE; t1_up := FALSE; 
    ELSIF ((x2 = FALSE) AND  ( TRUE ) AND  (x10 = TRUE) AND  (t0.Q = FALSE) AND  (t1.Q = FALSE)) THEN 
        cstate64 := 19; y2 := FALSE; y3 := FALSE; t0_start := FALSE;t1_start := FALSE; 
    ELSIF ((x2 = FALSE) AND  ( TRUE ) AND  (x10 = TRUE) AND  (t0.Q = FALSE) AND  (t1.Q = TRUE)) THEN 
        cstate64 := 20; y2 := FALSE; y3 := FALSE; t0_start := FALSE;t1_start := FALSE; 
    ELSIF ((x2 = FALSE) AND  ( TRUE ) AND  (x10 = TRUE) AND  (t0.Q = TRUE) AND  (t1.Q = FALSE)) THEN 
        cstate64 := 34; y2 := FALSE; y3 := FALSE; t0_start := FALSE;t1_start := FALSE; 
    ELSIF ((x2 = FALSE) AND  ( TRUE ) AND  (x10 = TRUE) AND  (t0.Q = TRUE) AND  (t1.Q = TRUE)) THEN 
        cstate64 := 33; y2 := FALSE; y3 := FALSE; t0_start := FALSE;t1_start := FALSE; 
    ELSIF ((x2 = TRUE) AND  ( TRUE ) AND  (x10 = FALSE) AND  (t0.Q = FALSE) AND  (t1.Q = FALSE)) THEN 
        cstate64 := 90; y2 := TRUE; y3 := TRUE; t0_start := FALSE;t1_start := FALSE; 
    ELSIF ((x2 = TRUE) AND  ( TRUE ) AND  (x10 = FALSE) AND  (t0.Q = FALSE) AND  (t1.Q = TRUE)) THEN 
        cstate64 := 84; y2 := TRUE; y3 := FALSE; t0_start := FALSE;t1_start := FALSE; 
    ELSIF ((x2 = TRUE) AND  ( TRUE ) AND  (x10 = FALSE) AND  (t0.Q = TRUE) AND  ( TRUE )) THEN 
        cstate64 := 69; y2 := FALSE; y3 := TRUE; t0_start := FALSE;t1_start := TRUE; t1_up := FALSE; 
    ELSIF ((x2 = TRUE) AND  ( TRUE ) AND  (x10 = TRUE) AND  (t0.Q = FALSE) AND  (t1.Q = FALSE)) THEN 
        cstate64 := 51; y2 := FALSE; y3 := FALSE; t0_start := FALSE;t1_start := FALSE; 
    ELSIF ((x2 = TRUE) AND  ( TRUE ) AND  (x10 = TRUE) AND  (t0.Q = FALSE) AND  (t1.Q = TRUE)) THEN 
        cstate64 := 52; y2 := FALSE; y3 := FALSE; t0_start := FALSE;t1_start := FALSE; 
    ELSIF ((x2 = TRUE) AND  ( TRUE ) AND  (x10 = TRUE) AND  (t0.Q = TRUE) AND  (t1.Q = FALSE)) THEN 
        cstate64 := 66; y2 := FALSE; y3 := FALSE; t0_start := FALSE;t1_start := FALSE; 
    ELSIF ((x2 = TRUE) AND  ( TRUE ) AND  (x10 = TRUE) AND  (t0.Q = TRUE) AND  (t1.Q = TRUE)) THEN 
        cstate64 := 65; y2 := FALSE; y3 := FALSE; t0_start := FALSE;t1_start := FALSE; 
    END_IF;
0:
    IF ((x2 = FALSE) AND  ( TRUE ) AND  (x10 = FALSE) AND  (t0.Q = FALSE) AND  (t1.Q = FALSE)) OR ((x2 = FALSE) AND  ( TRUE ) AND  (x10 = TRUE) AND  (t0.Q = FALSE) AND  ( TRUE )) THEN 
        cstate64 := 36; y2 := FALSE; y3 := FALSE; t0_start := FALSE;t1_start := FALSE; 
    ELSIF ((x2 = FALSE) AND  ( TRUE ) AND  (x10 = FALSE) AND  (t0.Q = FALSE) AND  (t1.Q = TRUE)) THEN 
        cstate64 := 36; y2 := FALSE; y3 := FALSE; t0_start := FALSE;t1_start := FALSE; 
    ELSIF ((x2 = FALSE) AND  ( TRUE ) AND  (x10 = FALSE) AND  (t0.Q = TRUE) AND  ( TRUE )) THEN 
        cstate64 := 33; y2 := FALSE; y3 := FALSE; t0_start := FALSE;t1_start := FALSE; 
    ELSIF ((x2 = FALSE) AND  ( TRUE ) AND  (x10 = TRUE) AND  (t0.Q = TRUE) AND  ( TRUE )) THEN 
        cstate64 := 33; y2 := FALSE; y3 := FALSE; t0_start := FALSE;t1_start := FALSE; 
    ELSIF ((x2 = TRUE) AND  ( TRUE ) AND  (x10 = FALSE) AND  (t0.Q = FALSE) AND  (t1.Q = FALSE)) OR ((x2 = TRUE) AND  ( TRUE ) AND  (x10 = TRUE) AND  (t0.Q = FALSE) AND  ( TRUE )) THEN 
        cstate64 := 68; y2 := FALSE; y3 := FALSE; t0_start := FALSE;t1_start := FALSE; 
    ELSIF ((x2 = TRUE) AND  ( TRUE ) AND  (x10 = FALSE) AND  (t0.Q = FALSE) AND  (t1.Q = TRUE)) THEN 
        cstate64 := 68; y2 := FALSE; y3 := FALSE; t0_start := FALSE;t1_start := FALSE; 
    ELSIF ((x2 = TRUE) AND  ( TRUE ) AND  ( TRUE ) AND  (t0.Q = TRUE) AND  ( TRUE )) THEN 
        cstate64 := 65; y2 := FALSE; y3 := FALSE; t0_start := FALSE;t1_start := FALSE; 
    END_IF;
51:
    IF ((x2 = FALSE) AND  ( TRUE ) AND  ( TRUE ) AND  (t0.Q = FALSE) AND  (t1.Q = FALSE)) THEN 
        cstate64 := 19; y2 := FALSE; y3 := FALSE; t0_start := FALSE;t1_start := FALSE; 
    ELSIF ((x2 = FALSE) AND  ( TRUE ) AND  (x10 = FALSE) AND  (t0.Q = FALSE) AND  (t1.Q = TRUE)) THEN 
        cstate64 := 20; y2 := FALSE; y3 := FALSE; t0_start := FALSE;t1_start := FALSE; 
    ELSIF ((x2 = FALSE) AND  ( TRUE ) AND  (x10 = FALSE) AND  (t0.Q = TRUE) AND  ( TRUE )) THEN 
        cstate64 := 37; y2 := FALSE; y3 := TRUE; t0_start := FALSE;t1_start := TRUE; t1_up := FALSE; 
    ELSIF ((x2 = FALSE) AND  ( TRUE ) AND  (x10 = TRUE) AND  (t0.Q = FALSE) AND  (t1.Q = TRUE)) THEN 
        cstate64 := 20; y2 := FALSE; y3 := FALSE; t0_start := FALSE;t1_start := FALSE; 
    ELSIF ((x2 = FALSE) AND  ( TRUE ) AND  (x10 = TRUE) AND  (t0.Q = TRUE) AND  (t1.Q = FALSE)) THEN 
        cstate64 := 34; y2 := FALSE; y3 := FALSE; t0_start := FALSE;t1_start := FALSE; 
    ELSIF ((x2 = FALSE) AND  ( TRUE ) AND  (x10 = TRUE) AND  (t0.Q = TRUE) AND  (t1.Q = TRUE)) THEN 
        cstate64 := 33; y2 := FALSE; y3 := FALSE; t0_start := FALSE;t1_start := FALSE; 
    ELSIF ((x2 = TRUE) AND  ( TRUE ) AND  ( TRUE ) AND  (t0.Q = FALSE) AND  (t1.Q = FALSE)) THEN 
        cstate64 := 51; y2 := FALSE; y3 := FALSE; t0_start := FALSE;t1_start := FALSE; 
    ELSIF ((x2 = TRUE) AND  ( TRUE ) AND  (x10 = FALSE) AND  (t0.Q = FALSE) AND  (t1.Q = TRUE)) THEN 
        cstate64 := 52; y2 := FALSE; y3 := FALSE; t0_start := FALSE;t1_start := FALSE; 
    ELSIF ((x2 = TRUE) AND  ( TRUE ) AND  (x10 = FALSE) AND  (t0.Q = TRUE) AND  ( TRUE )) THEN 
        cstate64 := 69; y2 := FALSE; y3 := TRUE; t0_start := FALSE;t1_start := TRUE; t1_up := FALSE; 
    ELSIF ((x2 = TRUE) AND  ( TRUE ) AND  (x10 = TRUE) AND  (t0.Q = FALSE) AND  (t1.Q = TRUE)) THEN 
        cstate64 := 52; y2 := FALSE; y3 := FALSE; t0_start := FALSE;t1_start := FALSE; 
    ELSIF ((x2 = TRUE) AND  ( TRUE ) AND  (x10 = TRUE) AND  (t0.Q = TRUE) AND  (t1.Q = FALSE)) THEN 
        cstate64 := 66; y2 := FALSE; y3 := FALSE; t0_start := FALSE;t1_start := FALSE; 
    ELSIF ((x2 = TRUE) AND  ( TRUE ) AND  (x10 = TRUE) AND  (t0.Q = TRUE) AND  (t1.Q = TRUE)) THEN 
        cstate64 := 65; y2 := FALSE; y3 := FALSE; t0_start := FALSE;t1_start := FALSE; 
    END_IF;
52:
    IF ((x2 = FALSE) AND  ( TRUE ) AND  (x10 = FALSE) AND  (t0.Q = FALSE) AND  (t1.Q = FALSE)) OR ((x2 = FALSE) AND  ( TRUE ) AND  (x10 = TRUE) AND  (t0.Q = FALSE) AND  ( TRUE )) THEN 
        cstate64 := 20; y2 := FALSE; y3 := FALSE; t0_start := FALSE;t1_start := FALSE; 
    ELSIF ((x2 = FALSE) AND  ( TRUE ) AND  (x10 = FALSE) AND  (t0.Q = FALSE) AND  (t1.Q = TRUE)) THEN 
        cstate64 := 20; y2 := FALSE; y3 := FALSE; t0_start := FALSE;t1_start := FALSE; 
    ELSIF ((x2 = FALSE) AND  ( TRUE ) AND  (x10 = FALSE) AND  (t0.Q = TRUE) AND  ( TRUE )) THEN 
        cstate64 := 40; y2 := FALSE; y3 := TRUE; t0_start := FALSE;t1_start := TRUE; t1_up := FALSE; 
    ELSIF ((x2 = FALSE) AND  ( TRUE ) AND  (x10 = TRUE) AND  (t0.Q = TRUE) AND  ( TRUE )) THEN 
        cstate64 := 33; y2 := FALSE; y3 := FALSE; t0_start := FALSE;t1_start := FALSE; 
    ELSIF ((x2 = TRUE) AND  ( TRUE ) AND  (x10 = FALSE) AND  (t0.Q = FALSE) AND  (t1.Q = FALSE)) OR ((x2 = TRUE) AND  ( TRUE ) AND  (x10 = TRUE) AND  (t0.Q = FALSE) AND  ( TRUE )) THEN 
        cstate64 := 52; y2 := FALSE; y3 := FALSE; t0_start := FALSE;t1_start := FALSE; 
    ELSIF ((x2 = TRUE) AND  ( TRUE ) AND  (x10 = FALSE) AND  (t0.Q = FALSE) AND  (t1.Q = TRUE)) THEN 
        cstate64 := 52; y2 := FALSE; y3 := FALSE; t0_start := FALSE;t1_start := FALSE; 
    ELSIF ((x2 = TRUE) AND  ( TRUE ) AND  (x10 = FALSE) AND  (t0.Q = TRUE) AND  ( TRUE )) THEN 
        cstate64 := 72; y2 := FALSE; y3 := TRUE; t0_start := FALSE;t1_start := TRUE; t1_up := FALSE; 
    ELSIF ((x2 = TRUE) AND  ( TRUE ) AND  (x10 = TRUE) AND  (t0.Q = TRUE) AND  ( TRUE )) THEN 
        cstate64 := 65; y2 := FALSE; y3 := FALSE; t0_start := FALSE;t1_start := FALSE; 
    END_IF;
72:
    IF ((x2 = FALSE) AND  ( TRUE ) AND  (x10 = FALSE) AND  (t0.Q = FALSE) AND  (t1.Q = FALSE)) THEN 
        cstate64 := 44; y2 := FALSE; y3 := TRUE; t0_start := FALSE;t1_start := FALSE; 
    ELSIF ((x2 = FALSE) AND  ( TRUE ) AND  (x10 = FALSE) AND  (t0.Q = FALSE) AND  (t1.Q = TRUE)) THEN 
        cstate64 := 36; y2 := FALSE; y3 := FALSE; t0_start := FALSE;t1_start := FALSE; 
    ELSIF ((x2 = FALSE) AND  ( TRUE ) AND  (x10 = FALSE) AND  (t0.Q = TRUE) AND  (t1.Q = FALSE)) THEN 
        cstate64 := 40; y2 := FALSE; y3 := TRUE; t0_start := FALSE;t1_start := FALSE; 
    ELSIF ((x2 = FALSE) AND  ( TRUE ) AND  (x10 = FALSE) AND  (t0.Q = TRUE) AND  (t1.Q = TRUE)) THEN 
        cstate64 := 33; y2 := FALSE; y3 := FALSE; t0_start := FALSE;t1_start := FALSE; 
    ELSIF ((x2 = FALSE) AND  ( TRUE ) AND  (x10 = TRUE) AND  (t0.Q = FALSE) AND  (t1.Q = FALSE)) THEN 
        cstate64 := 35; y2 := FALSE; y3 := FALSE; t0_start := FALSE;t1_start := FALSE; 
    ELSIF ((x2 = FALSE) AND  ( TRUE ) AND  (x10 = TRUE) AND  (t0.Q = FALSE) AND  (t1.Q = TRUE)) THEN 
        cstate64 := 36; y2 := FALSE; y3 := FALSE; t0_start := FALSE;t1_start := FALSE; 
    ELSIF ((x2 = FALSE) AND  ( TRUE ) AND  (x10 = TRUE) AND  (t0.Q = TRUE) AND  (t1.Q = FALSE)) THEN 
        cstate64 := 34; y2 := FALSE; y3 := FALSE; t0_start := FALSE;t1_start := FALSE; 
    ELSIF ((x2 = FALSE) AND  ( TRUE ) AND  (x10 = TRUE) AND  (t0.Q = TRUE) AND  (t1.Q = TRUE)) THEN 
        cstate64 := 33; y2 := FALSE; y3 := FALSE; t0_start := FALSE;t1_start := FALSE; 
    ELSIF ((x2 = TRUE) AND  ( TRUE ) AND  (x10 = FALSE) AND  (t0.Q = FALSE) AND  (t1.Q = FALSE)) THEN 
        cstate64 := 76; y2 := FALSE; y3 := TRUE; t0_start := FALSE;t1_start := FALSE; 
    ELSIF ((x2 = TRUE) AND  ( TRUE ) AND  (x10 = FALSE) AND  (t0.Q = FALSE) AND  (t1.Q = TRUE)) THEN 
        cstate64 := 68; y2 := FALSE; y3 := FALSE; t0_start := FALSE;t1_start := FALSE; 
    ELSIF ((x2 = TRUE) AND  ( TRUE ) AND  (x10 = FALSE) AND  (t0.Q = TRUE) AND  (t1.Q = FALSE)) THEN 
        cstate64 := 72; y2 := FALSE; y3 := TRUE; t0_start := FALSE;t1_start := FALSE; 
    ELSIF ((x2 = TRUE) AND  ( TRUE ) AND  ( TRUE ) AND  (t0.Q = TRUE) AND  (t1.Q = TRUE)) THEN 
        cstate64 := 65; y2 := FALSE; y3 := FALSE; t0_start := FALSE;t1_start := FALSE; 
    ELSIF ((x2 = TRUE) AND  ( TRUE ) AND  (x10 = TRUE) AND  (t0.Q = FALSE) AND  (t1.Q = FALSE)) THEN 
        cstate64 := 67; y2 := FALSE; y3 := FALSE; t0_start := FALSE;t1_start := FALSE; 
    ELSIF ((x2 = TRUE) AND  ( TRUE ) AND  (x10 = TRUE) AND  (t0.Q = FALSE) AND  (t1.Q = TRUE)) THEN 
        cstate64 := 68; y2 := FALSE; y3 := FALSE; t0_start := FALSE;t1_start := FALSE; 
    ELSIF ((x2 = TRUE) AND  ( TRUE ) AND  (x10 = TRUE) AND  (t0.Q = TRUE) AND  (t1.Q = FALSE)) THEN 
        cstate64 := 66; y2 := FALSE; y3 := FALSE; t0_start := FALSE;t1_start := FALSE; 
    END_IF;
73:
    IF ((x2 = FALSE) AND  ( TRUE ) AND  (x10 = FALSE) AND  (t0.Q = FALSE) AND  (t1.Q = FALSE)) THEN 
        cstate64 := 41; y2 := FALSE; y3 := TRUE; t0_start := FALSE;t1_start := FALSE; 
    ELSIF ((x2 = FALSE) AND  ( TRUE ) AND  (x10 = FALSE) AND  (t0.Q = FALSE) AND  (t1.Q = TRUE)) THEN 
        cstate64 := 36; y2 := FALSE; y3 := FALSE; t0_start := FALSE;t1_start := FALSE; 
    ELSIF ((x2 = FALSE) AND  ( TRUE ) AND  (x10 = FALSE) AND  (t0.Q = TRUE) AND  ( TRUE )) THEN 
        cstate64 := 37; y2 := FALSE; y3 := TRUE; t0_start := FALSE;t1_start := TRUE; t1_up := FALSE; 
    ELSIF ((x2 = FALSE) AND  ( TRUE ) AND  (x10 = TRUE) AND  (t0.Q = FALSE) AND  (t1.Q = FALSE)) THEN 
        cstate64 := 35; y2 := FALSE; y3 := FALSE; t0_start := FALSE;t1_start := FALSE; 
    ELSIF ((x2 = FALSE) AND  ( TRUE ) AND  (x10 = TRUE) AND  (t0.Q = FALSE) AND  (t1.Q = TRUE)) THEN 
        cstate64 := 36; y2 := FALSE; y3 := FALSE; t0_start := FALSE;t1_start := FALSE; 
    ELSIF ((x2 = FALSE) AND  ( TRUE ) AND  (x10 = TRUE) AND  (t0.Q = TRUE) AND  (t1.Q = FALSE)) THEN 
        cstate64 := 34; y2 := FALSE; y3 := FALSE; t0_start := FALSE;t1_start := FALSE; 
    ELSIF ((x2 = FALSE) AND  ( TRUE ) AND  (x10 = TRUE) AND  (t0.Q = TRUE) AND  (t1.Q = TRUE)) THEN 
        cstate64 := 33; y2 := FALSE; y3 := FALSE; t0_start := FALSE;t1_start := FALSE; 
    ELSIF ((x2 = TRUE) AND  ( TRUE ) AND  (x10 = FALSE) AND  (t0.Q = FALSE) AND  (t1.Q = FALSE)) THEN 
        cstate64 := 73; y2 := FALSE; y3 := TRUE; t0_start := FALSE;t1_start := FALSE; 
    ELSIF ((x2 = TRUE) AND  ( TRUE ) AND  (x10 = FALSE) AND  (t0.Q = FALSE) AND  (t1.Q = TRUE)) THEN 
        cstate64 := 68; y2 := FALSE; y3 := FALSE; t0_start := FALSE;t1_start := FALSE; 
    ELSIF ((x2 = TRUE) AND  ( TRUE ) AND  (x10 = FALSE) AND  (t0.Q = TRUE) AND  ( TRUE )) THEN 
        cstate64 := 69; y2 := FALSE; y3 := TRUE; t0_start := FALSE;t1_start := TRUE; t1_up := FALSE; 
    ELSIF ((x2 = TRUE) AND  ( TRUE ) AND  (x10 = TRUE) AND  (t0.Q = FALSE) AND  (t1.Q = FALSE)) THEN 
        cstate64 := 67; y2 := FALSE; y3 := FALSE; t0_start := FALSE;t1_start := FALSE; 
    ELSIF ((x2 = TRUE) AND  ( TRUE ) AND  (x10 = TRUE) AND  (t0.Q = FALSE) AND  (t1.Q = TRUE)) THEN 
        cstate64 := 68; y2 := FALSE; y3 := FALSE; t0_start := FALSE;t1_start := FALSE; 
    ELSIF ((x2 = TRUE) AND  ( TRUE ) AND  (x10 = TRUE) AND  (t0.Q = TRUE) AND  (t1.Q = FALSE)) THEN 
        cstate64 := 66; y2 := FALSE; y3 := FALSE; t0_start := FALSE;t1_start := FALSE; 
    ELSIF ((x2 = TRUE) AND  ( TRUE ) AND  (x10 = TRUE) AND  (t0.Q = TRUE) AND  (t1.Q = TRUE)) THEN 
        cstate64 := 65; y2 := FALSE; y3 := FALSE; t0_start := FALSE;t1_start := FALSE; 
    END_IF;
76:
    IF ((x2 = FALSE) AND  ( TRUE ) AND  (x10 = FALSE) AND  (t0.Q = FALSE) AND  (t1.Q = FALSE)) THEN 
        cstate64 := 44; y2 := FALSE; y3 := TRUE; t0_start := FALSE;t1_start := FALSE; 
    ELSIF ((x2 = FALSE) AND  ( TRUE ) AND  (x10 = FALSE) AND  (t0.Q = FALSE) AND  (t1.Q = TRUE)) THEN 
        cstate64 := 36; y2 := FALSE; y3 := FALSE; t0_start := FALSE;t1_start := FALSE; 
    ELSIF ((x2 = FALSE) AND  ( TRUE ) AND  (x10 = FALSE) AND  (t0.Q = TRUE) AND  (t1.Q = FALSE)) THEN 
        cstate64 := 40; y2 := FALSE; y3 := TRUE; t0_start := FALSE;t1_start := TRUE; t1_up := FALSE; 
    ELSIF ((x2 = FALSE) AND  ( TRUE ) AND  (x10 = FALSE) AND  (t0.Q = TRUE) AND  (t1.Q = TRUE)) THEN 
        cstate64 := 37; y2 := FALSE; y3 := TRUE; t0_start := FALSE;t1_start := TRUE; t1_up := FALSE; 
    ELSIF ((x2 = FALSE) AND  ( TRUE ) AND  (x10 = TRUE) AND  (t0.Q = FALSE) AND  (t1.Q = FALSE)) THEN 
        cstate64 := 35; y2 := FALSE; y3 := FALSE; t0_start := FALSE;t1_start := FALSE; 
    ELSIF ((x2 = FALSE) AND  ( TRUE ) AND  (x10 = TRUE) AND  (t0.Q = FALSE) AND  (t1.Q = TRUE)) THEN 
        cstate64 := 36; y2 := FALSE; y3 := FALSE; t0_start := FALSE;t1_start := FALSE; 
    ELSIF ((x2 = FALSE) AND  ( TRUE ) AND  (x10 = TRUE) AND  (t0.Q = TRUE) AND  (t1.Q = FALSE)) THEN 
        cstate64 := 34; y2 := FALSE; y3 := FALSE; t0_start := FALSE;t1_start := FALSE; 
    ELSIF ((x2 = FALSE) AND  ( TRUE ) AND  (x10 = TRUE) AND  (t0.Q = TRUE) AND  (t1.Q = TRUE)) THEN 
        cstate64 := 33; y2 := FALSE; y3 := FALSE; t0_start := FALSE;t1_start := FALSE; 
    ELSIF ((x2 = TRUE) AND  ( TRUE ) AND  (x10 = FALSE) AND  (t0.Q = FALSE) AND  (t1.Q = FALSE)) THEN 
        cstate64 := 76; y2 := FALSE; y3 := TRUE; t0_start := FALSE;t1_start := FALSE; 
    ELSIF ((x2 = TRUE) AND  ( TRUE ) AND  (x10 = FALSE) AND  (t0.Q = FALSE) AND  (t1.Q = TRUE)) THEN 
        cstate64 := 68; y2 := FALSE; y3 := FALSE; t0_start := FALSE;t1_start := FALSE; 
    ELSIF ((x2 = TRUE) AND  ( TRUE ) AND  (x10 = FALSE) AND  (t0.Q = TRUE) AND  (t1.Q = FALSE)) THEN 
        cstate64 := 72; y2 := FALSE; y3 := TRUE; t0_start := FALSE;t1_start := TRUE; t1_up := FALSE; 
    ELSIF ((x2 = TRUE) AND  ( TRUE ) AND  (x10 = FALSE) AND  (t0.Q = TRUE) AND  (t1.Q = TRUE)) THEN 
        cstate64 := 69; y2 := FALSE; y3 := TRUE; t0_start := FALSE;t1_start := TRUE; t1_up := FALSE; 
    ELSIF ((x2 = TRUE) AND  ( TRUE ) AND  (x10 = TRUE) AND  (t0.Q = FALSE) AND  (t1.Q = FALSE)) THEN 
        cstate64 := 67; y2 := FALSE; y3 := FALSE; t0_start := FALSE;t1_start := FALSE; 
    ELSIF ((x2 = TRUE) AND  ( TRUE ) AND  (x10 = TRUE) AND  (t0.Q = FALSE) AND  (t1.Q = TRUE)) THEN 
        cstate64 := 68; y2 := FALSE; y3 := FALSE; t0_start := FALSE;t1_start := FALSE; 
    ELSIF ((x2 = TRUE) AND  ( TRUE ) AND  (x10 = TRUE) AND  (t0.Q = TRUE) AND  (t1.Q = FALSE)) THEN 
        cstate64 := 66; y2 := FALSE; y3 := FALSE; t0_start := FALSE;t1_start := FALSE; 
    ELSIF ((x2 = TRUE) AND  ( TRUE ) AND  (x10 = TRUE) AND  (t0.Q = TRUE) AND  (t1.Q = TRUE)) THEN 
        cstate64 := 65; y2 := FALSE; y3 := FALSE; t0_start := FALSE;t1_start := FALSE; 
    END_IF;
END_CASE;

